(* IEC 61131-3 sources: plcassist-cli/packages/volt-lsp-iec/test-corpus/pro2193/Device/Plc Logic/Application/09 Misc/Library Manager/L_MC4P_RoboticHandling (part 3) *)

(* ---- L_MC4P_PATHREFFROMFILE.fb ---- *)
FUNCTION_BLOCK L_MC4P_PATHREFFROMFILE
VAR_INPUT
	XEXECUTE : BOOL;
	SFILENAME : STRING;
	XABORT : BOOL;
	DWSKIPMASK : DWORD := 0;
	LIBLOCKSEARCHLINENO : LINT := 0;
END_VAR
VAR_OUTPUT
	XDONE : BOOL;
	XBUSY : BOOL;
	XCOMMANDABORTED : BOOL;
	XERROR : BOOL;
	EERRORID : L_IE1P_Error;
	XDECODING : BOOL;
	LILINENODECODED : LINT;
	SLINEDECODED : STRING;
END_VAR
VAR
	LIBLOCKSEARCHLINENO_INT : LINT;
	IFILENO_INT : INT;
	XINTERPRETERHALT_INT : BOOL;
	XMOVEPATHACTIVE_INT : BOOL;
	WACTIVEMFUNCTION_INT : WORD;
	LISOURCELINENO_INT : LINT;
	XABORTACTIVE : BOOL;
	_XDONE : BOOL;
	_XBUSY : BOOL;
	_XCOMMANDABORTED : BOOL;
	_XDECODING : BOOL;
	SFILEADRESS : STRING;
	ITACKEDNUMOFELEMENTSINCYCLE_INT : INT := 0;
	IDECODEMAXNUMOFELEMENTS_INT : INT := 2;
	IDECODEMAXNUMOFELEMENTSFIRSTTIME_INT : INT := 3;
	IDECODENUMOFELEMENTS_INT : INT;
	FB_DECODENCPROGDATA : L_MC1P_StackControlArray := STRUCT(iMaxLegth := GVL_MovePath.gciNumOfPathFiles);
	SCHEADDATA : L_MC4P_AsciiDecoderHeadData;
	RSCACTFILEDATA : REFERENCE TO L_MC4P_AsciiDecoderFileData;
	XHALTATMOS_INT : BOOL := TRUE;
	XIGNOREMCOMMANDS_INT : BOOL;
	XNEWFILE_INT : BOOL;
	LRCIRCLTARGETTOLERANCE_INT : LREAL := 0.1;
	FB_SEMA : L_MC1P_CriticalSection;
	ITAKEELEMENTCNT : INT;
	IADDELEMENTCNT : INT;
	FB_DECODEMOVEDATALOWTASK : L_MC1P_StackControlArray := STRUCT(iMaxLegth := GVL_MovePath.gciNumOfDecodeAsciiData);
	FB_DECODEMOVEDATAMOTIONTASK : L_MC1P_StackControlArray := STRUCT(iMaxLegth := GVL_MovePath.gciNumOfDecodeAsciiData);
	ASCDECODEMOVEDATA_INT : ARRAY [1..GVL_MovePath.gciNumOfDecodeAsciiData] OF L_MC4P_Parameter_MCMove;
	IELEMENINARRAYDECODING : INT;
	FB_DECODEMOVEDATALOWTASK_RESERVE : L_MC1P_StackControlArray := STRUCT(iMaxLegth := GVL_MovePath.gciNumOfDecodeAsciiData_reserve);
	ASCDECODEMOVEDATA_RESERVE : ARRAY [1..GVL_MovePath.gciNumOfDecodeAsciiData_reserve] OF L_MC4P_Parameter_MCMove;
	XERROR_DECODERENDLOOP : BOOL;
	DWTIMEOUTCNT : DWORD := 0;
	DWTIMEOUT : DWORD := 100000;
	XERROR_TIMEOUT : BOOL;
	DWTIMEOUT_MASK : DWORD;
	WTIMEOUTDECODERSTATE : WORD;
	WSTATE : WORD;
	XID1 : BOOL;
	XWID_INT : POINTER TO BOOL := ADR(xId1);
	XSETPATHDATAACTIVE_INT : BOOL;
	XSETPATHDATAACTIVE_OLD : BOOL;
	REQUESTSINFO : DWORD;
	REQUESTSINFO_OLD : DWORD;
	DWRTRIG : DWORD;
	DWFTRIG : DWORD;
	XRESETOUTPUTS : BOOL;
	XERROR_INVALIDSYNCDATA : BOOL;
	BYERRORADRESS : BYTE;
	STERRORADRESSVALUE : STRING;
	XPATHREFABORT : BOOL;
	XDECODEINNEXTTASKCYCLE : BOOL;
	XFBISABORTED : BOOL;
	SFILE_INT : STRING := '';
	XDECODEBUSY_INT : BOOL;
	XDECODEDONE_INT : BOOL;
	XDECODEERROR_INT : BOOL;
	EDECODEEERRORID_INT : L_IE1P_Error;
	DWINTERNALID_INT : DWORD;
	STDECODEERRORLINE : STRING;
	RES : SYSFILE.RTS_IEC_RESULT;
	HFILE : SYSFILE.RTS_IEC_HANDLE;
	UDILENGTHFILE : UDINT;
	XTESTINMOTIONTASK : BOOL := FALSE;
	EXCEPTIONCODE : __SYSTEM.ExceptionCode;
	DWPREDECODERIDLECYCLES : DWORD := 0;
	DWPOSTDECODERIDLECYCLES : DWORD := 0;
	BLOCKSEARCHENABLED : BOOL;
	DATATYPE : WORD;
	DWTIMEOUTMASK : DWORD;
	ENDELEMENT : POINTER TO L_MC4P_Parameter_MCMove;
	ENDIDX : INT;
	POSTDECODERIDLECYCLES : DWORD;
	PREDECODERIDLECYCLES : DWORD;
	SETCIRCTARGETTOLERANCE : LREAL;
	SIZE : UDINT;
	STARTELEMENT : POINTER TO L_MC4P_Parameter_MCMove;
	STARTIDX : INT;
	STERRORCOMMAND : STRING;
	TAKEELEMENT : POINTER TO L_MC4P_Parameter_MCMove;
	XDECODEINMOTIONTASK : BOOL;
	XHALTATMOS : BOOL;
	XIGNOREMCOMMANDS : BOOL;
	XINTERPRETERHALT : BOOL;
END_VAR
END_FUNCTION_BLOCK

METHOD ABORTFB
END_METHOD

METHOD CALL_ALLOCPOINTADR
END_METHOD

METHOD CALL_ERRORHANDLER
END_METHOD

METHOD CALL_FBMETHODS
END_METHOD

METHOD CALL_OUTPUT
END_METHOD

METHOD CALL_REQUESTS_EXT
END_METHOD

METHOD CALL_RESETCOMMANDS
END_METHOD

METHOD CALL_RESETOUTPUT
END_METHOD

METHOD CALL_RESETSTATUS
END_METHOD

METHOD CALL_STATEMACHINE
END_METHOD

METHOD CALL_SYNCDECODEMOVEDATA
END_METHOD

METHOD FUN_DECODEAUX : BOOL
VAR_IN_OUT
	STADRESSVALUE : STRING(255);
	SCDECODEHEADDATA : L_MC4P_AsciiDecoderHeadData;
END_VAR
END_METHOD

METHOD FUN_DECODEADRESS : BOOL
VAR_OUTPUT
	XERROR : BOOL;
	EERRORID : L_IE1P_Error;
END_VAR
VAR_IN_OUT
	BYADRESS : BYTE;
	STADRESSVALUE : STRING(255);
	SCDECODEHEADDATA : L_MC4P_AsciiDecoderHeadData;
END_VAR
END_METHOD

METHOD FUN_DECODEG : BOOL
VAR_IN_OUT
	LIADRESSVALUE : LINT;
	SCDECODEHEADDATA : L_MC4P_AsciiDecoderHeadData;
END_VAR
END_METHOD

METHOD FUN_DECODEGOTO : BOOL
VAR_OUTPUT
	XERROR : BOOL;
	EERRORID : L_IE1P_Error;
END_VAR
VAR_IN_OUT
	STADRESSVALUE : STRING(255);
	SCDECODEHEADDATA : L_MC4P_AsciiDecoderHeadData;
END_VAR
END_METHOD

METHOD FUN_DECODEH : BOOL
VAR_IN_OUT
	STADRESSVALUE : STRING(255);
	SCDECODEHEADDATA : L_MC4P_AsciiDecoderHeadData;
	XERROR : BOOL;
	EERRORID : L_IE1P_Error;
END_VAR
END_METHOD

METHOD FUN_DECODEI : BOOL
VAR_IN_OUT
	STADRESSVALUE : STRING(255);
	SCDECODEHEADDATA : L_MC4P_AsciiDecoderHeadData;
END_VAR
END_METHOD

METHOD FUN_DECODEIFCASE : BOOL
VAR_INPUT
	STLINE : STRING(255);
END_VAR
VAR_OUTPUT
	XERROR : BOOL;
	EERRORID : L_IE1P_Error;
END_VAR
VAR_IN_OUT
	SCDECODEHEADDATA : L_MC4P_AsciiDecoderHeadData;
END_VAR
END_METHOD

METHOD FUN_DECODEL : BOOL
VAR_IN_OUT
	STADRESSVALUE : STRING(255);
	SCDECODEHEADDATA : L_MC4P_AsciiDecoderHeadData;
	XERROR : BOOL;
	EERRORID : L_IE1P_Error;
END_VAR
END_METHOD

METHOD FUN_DECODELINE : BOOL
VAR_OUTPUT
	XGETNEXTSOURCELINE : BOOL;
	XELEMENTDECODED : BOOL;
	XERROR : BOOL;
	EERRORID : L_IE1P_Error;
END_VAR
VAR_IN_OUT
	SCDECODEHEADDATA : L_MC4P_AsciiDecoderHeadData;
	SCDECODEMOVEDATA : L_MC4P_Parameter_MCMove;
END_VAR
END_METHOD

METHOD FUN_DECODEM : BOOL
VAR_IN_OUT
	LIADRESSVALUE : LINT;
	SCDECODEHEADDATA : L_MC4P_AsciiDecoderHeadData;
	XERROR : BOOL;
	EERRORID : L_IE1P_Error;
END_VAR
END_METHOD

METHOD FUN_DECODEN : BOOL
VAR_IN_OUT
	STADRESSVALUE : STRING(255);
	SCDECODEHEADDATA : L_MC4P_AsciiDecoderHeadData;
END_VAR
END_METHOD

METHOD FUN_DECODEO : BOOL
VAR_IN_OUT
	STADRESSVALUE : STRING(255);
	SCDECODEHEADDATA : L_MC4P_AsciiDecoderHeadData;
	XERROR : BOOL;
	EERRORID : L_IE1P_Error;
END_VAR
END_METHOD

METHOD FUN_DECODEP : BOOL
VAR_IN_OUT
	STADRESSVALUE : STRING(255);
	SCDECODEHEADDATA : L_MC4P_AsciiDecoderHeadData;
END_VAR
END_METHOD

METHOD FUN_DELETECOMMENTS : BOOL
VAR_OUTPUT
	STCOMMENT : STRING;
	ILINESIZE : INT;
END_VAR
VAR_IN_OUT
	STLINE : STRING(255);
END_VAR
END_METHOD

METHOD FUN_DELETECOMMENTS_TYPE1 : BOOL
VAR_IN_OUT
	STLINE : STRING(255);
	STCOMMENT : STRING;
	ICOMMENTPOS : INT;
END_VAR
END_METHOD

METHOD FUN_DELETECOMMENTS_TYPE2 : BOOL
VAR_INPUT
	ICOMMENTTYPE : INT;
END_VAR
VAR_IN_OUT
	STLINE : STRING(255);
	STCOMMENT : STRING;
END_VAR
END_METHOD

METHOD FUN_FINDJUMPTARB : BOOL
VAR_INPUT
	LIJUMPTARGET : LINT;
	UDIFILELENGTH : UDINT;
	UDIPOS : UDINT;
	UDIPOSSTART : UDINT;
END_VAR
VAR_OUTPUT
	UDITARLINEPOS : UDINT;
	XERROR : BOOL;
	EERRORID : L_IE1P_Error;
END_VAR
END_METHOD

METHOD FUN_FINDJUMPTARF : BOOL
VAR_INPUT
	LIJUMPTARGET : LINT;
	UDIFILELENGTH : UDINT;
	UDIPOS : UDINT;
END_VAR
VAR_OUTPUT
	UDITARLINEPOS : UDINT;
	XERROR : BOOL;
	EERRORID : L_IE1P_Error;
END_VAR
END_METHOD

METHOD FUN_GOTO : BOOL
VAR_OUTPUT
	XERROR : BOOL;
	EERRORID : L_IE1P_Error;
END_VAR
VAR_IN_OUT
	SCDECODEHEADDATA : L_MC4P_AsciiDecoderHeadData;
	STLINE : STRING(255);
END_VAR
END_METHOD

METHOD FUN_GETADRESS : BOOL
VAR_OUTPUT
	ILINESIZE : INT;
	BYADRESS : BYTE;
	SADRESSVALUE : STRING;
END_VAR
VAR_IN_OUT
	STLINE : STRING(255);
END_VAR
END_METHOD

METHOD FUN_ISALPHACHAR : BOOL
VAR_INPUT
	BYCHAR : BYTE;
END_VAR
END_METHOD

METHOD FUN_READLINE : L_IE1P_Error
VAR_INPUT
	UDIPOSIN : UDINT;
	XEXITCLOSEFILE : BOOL;
	XFINDSTARTCOMAND : BOOL;
END_VAR
VAR_OUTPUT
	UDIPOSOUT : UDINT;
	ILINESIZE : INT;
	IPOSLF : INT;
	IPOSNL : INT;
	UDIRESULTFILEOPEN : UDINT;
	UDIRESULTREADSTRING : UDINT;
	XENDOFFILE : BOOL;
	XLASTLINE : BOOL;
	XSTART : BOOL;
END_VAR
VAR_IN_OUT
	HFILE : SYSFILE.RTS_IEC_HANDLE;
	RES : SYSFILE.RTS_IEC_ResULT;
	STLINE : STRING(255);
END_VAR
END_METHOD

METHOD FUN_READLINEBACK : BOOL
VAR_INPUT
	UDIPOSIN : UDINT;
	XEXITCLOSEFILE : BOOL;
	UDIPOSSTART : UDINT := 0;
END_VAR
VAR_OUTPUT
	UDIPOSOUT : UDINT;
	ILINESIZE : INT;
	UDIRESULTFILEOPEN : UDINT;
	XSTARTOFFILE : BOOL;
END_VAR
VAR_IN_OUT
	HFILE : SYSFILE.RTS_IEC_HANDLE;
	RES : SYSFILE.RTS_IEC_ResULT;
	STLINE : STRING(255);
END_VAR
END_METHOD

METHOD FUN_REPLACEVAR : BOOL
VAR_IN_OUT
	STVALUE : STRING(255);
END_VAR
END_METHOD

METHOD FUN_STRING_PLCVARIABLE_TO_LINT : BOOL
VAR_INPUT
	STVALUE : STRING(255);
END_VAR
VAR_OUTPUT
	LIVALUE : LINT;
END_VAR
END_METHOD

METHOD FUN_STRING_PLCVARIABLE_TO_LREAL : BOOL
VAR_INPUT
	STVALUE : STRING(255);
END_VAR
VAR_OUTPUT
	LRVALUE : LREAL;
END_VAR
END_METHOD

METHOD FUN_STRING_TO_LINT : BOOL
VAR_INPUT
	STVALUE : STRING;
	XVARALLOWED : BOOL;
END_VAR
VAR_OUTPUT
	LIVALUE : LINT;
END_VAR
END_METHOD

METHOD FUN_STRING_TO_LREAL : BOOL
VAR_INPUT
	STVALUE : STRING(255);
END_VAR
VAR_OUTPUT
	LRVALUE : LREAL;
END_VAR
END_METHOD

METHOD FUN_SHUNTINGYARD : BOOL
VAR_INPUT
	STVALUE : STRING(255);
END_VAR
VAR_OUTPUT
	SCVALUE : L_UBUP_Variable;
END_VAR
END_METHOD

METHOD CALL_DECODER
END_METHOD

METHOD CALL_DECODER_READASCIIFILE
END_METHOD

METHOD EXECUTEFREERUNTASK
END_METHOD

METHOD FUN_CLOSEFILE
END_METHOD

METHOD INIT_HEADDATA
VAR_IN_OUT
	SCDECODEHEADDATA : L_MC4P_AsciiDecoderHeadData;
END_VAR
END_METHOD

METHOD MAIN
END_METHOD

METHOD GETID : __XWORD
END_METHOD

METHOD GETPATHDATA : ARRAY [1..GVL_MovePath.gciNumOfDecodeAsciiData] OF POINTER TO L_MC4P_Parameter_MCMove
END_METHOD

METHOD GETPATHDATAACTIVE : BOOL
END_METHOD

METHOD GETSTATUS : DWORD
END_METHOD

METHOD SETABORT
END_METHOD

METHOD SETACTIVEMFUNCTION
VAR_INPUT
	WACTIVEMFUNCTION : WORD;
END_VAR
END_METHOD

METHOD SETMOVEPATHACTIVE
VAR_INPUT
	XMOVEPATHACTIVE : BOOL;
END_VAR
END_METHOD

METHOD SETPATHDATAACTIVE
VAR_INPUT
	XPATHDATAACTIVE : BOOL;
END_VAR
END_METHOD

METHOD CALL_INIT
END_METHOD

METHOD CALL_S000_CYCLIC
END_METHOD

METHOD ABORT : UDINT
END_METHOD

METHOD EXECUTE : UDINT
END_METHOD

(* ---- L_MC4P_PATHREFMONITOR.fb ---- *)
FUNCTION_BLOCK L_MC4P_PATHREFMONITOR
VAR_INPUT
	XEXECUTE : BOOL;
	XABORT : BOOL;
	ITFPATHREF : MC_PATH_REF;
	SCSKIP : L_MC4P_SkipGCode;
	ASCDATA : POINTER TO L_MC4P_PathRefMonitorData;
END_VAR
VAR_OUTPUT
	XDONE : BOOL;
	XBUSY : BOOL;
	XCOMMANDABORTED : BOOL;
	XERROR : BOOL;
	EERRORID : L_IE1P_Error;
	UDINEWESTELEMENT : UDINT;
	UDIELEMENTCOUNT : UDINT;
END_VAR
VAR
	_ITFPATHREF : MC_PATH_REF;
	_UDISTARTIDX : UDINT;
	_UDIENDIDX : UDINT;
	_UDIREADIDX : UDINT;
	_UDILOWER : UDINT;
	_UDIUPPER : UDINT;
	_UDISIZE : UDINT;
	_DWSTATUS : DWORD;
	_XREINIT : BOOL := FALSE;
	_XDATADIALOG : BOOL := FALSE;
	_UDIVISUARRIDX : UDINT := 0;
	_PSCDATAARR : POINTER TO L_MC4P_PathRefMonitorData;
	_PSCDATAVISU : POINTER TO L_MC4P_PathRefMonitorData;
	_SCDATAINITIAL : L_MC4P_PathRefMonitorData;
	_ISKIPVIEWFRAME : INT := 0;
	_MODEL : L_UBUP_BehaviourModel_ETrigA;
END_VAR
END_FUNCTION_BLOCK

METHOD MAPOUTPUTS
END_METHOD

METHOD CYCLICACTION
VAR_INPUT
	ITFTIMINGCONTROLLER : L_UBUP.L_UBUP_ITimingController;
END_VAR
VAR_OUTPUT
	XCOMPLETE : BOOL;
	XABORT : BOOL;
	IERRORID : INT;
END_VAR
END_METHOD

METHOD FINALIZEACTION
VAR_INPUT
	XABORTPROPOSED : BOOL;
	IERRORIDPROPOSED : INT;
END_VAR
VAR_OUTPUT
	XCOMPLETE : BOOL;
	XABORT : BOOL;
	IERRORID : INT;
END_VAR
END_METHOD

METHOD RESETACTION
VAR_OUTPUT
	XCOMPLETE : BOOL;
END_VAR
END_METHOD

METHOD STARTACTION
VAR_OUTPUT
	XCOMPLETE : BOOL;
	IERRORID : INT;
END_VAR
END_METHOD

METHOD FB_INIT : BOOL
VAR_INPUT
	BINITRETAINS : BOOL;
	BINCOPYCODE : BOOL;
END_VAR
END_METHOD

METHOD APPENDDATASET : BOOL
VAR_INPUT
	PMCMOVE : POINTER TO L_MC4P_Parameter_MCMove;
END_VAR
END_METHOD

METHOD SKIP : BOOL
VAR_INPUT
	PMCMOVE : POINTER TO L_MC4P_Parameter_MCMove;
END_VAR
END_METHOD

(* ---- L_MC4P_PICKANDPLACEMEMORY.fb ---- *)
FUNCTION_BLOCK L_MC4P_PICKANDPLACEMEMORY
VAR_INPUT
	FB_SEMAMOVEFBS : L_MC1P_CriticalSection;
	AMC_MOVELINREL : ARRAY [1..3] OF L_MC4P_MoveLinearRelative_Internal;
	AFB_MOVEELLIPTICAL : ARRAY [1..3] OF L_MC4P_MoveEllipticalAbsolutePnP_Internal;
	AFB_MOVESPLINE : ARRAY [1..3] OF L_MC4P_MoveSplinePnP_Internal;
	AMC_MOVELINABS1 : ARRAY [1..10] OF L_MC4P_MoveLinearAbsolute_Internal;
	AMC_MOVELINABS2 : ARRAY [1..10] OF L_MC4P_MoveLinearAbsolute_Internal;
	AMC_MOVELINABS3 : ARRAY [1..10] OF L_MC4P_MoveLinearAbsolute_Internal;
	AMC_MOVELINABS4 : ARRAY [1..3] OF L_MC4P_MoveLinearAbsolute_Internal;
	AMC_MOVELINABS5 : ARRAY [1..2] OF L_MC4P_MoveLinearAbsolute_Internal;
	AMC_MOVEDIRABS1 : ARRAY [1..10] OF L_MC4P_MoveDirectAbsolute_Internal;
	AMC_MOVEDIRABS2 : ARRAY [1..10] OF L_MC4P_MoveDirectAbsolute_Internal;
	AMC_MOVEDIRREL : ARRAY [1..1] OF L_MC4P_MoveDirectRelative_Internal;
	AFB_GROUPWAITTIME : ARRAY [1..3] OF L_MC4P_GroupWaitTime_Internal;
	ASCPROFILEPARMEM : ARRAY [1..10] OF ARRAY [1..10] OF L_MC4P_scPickAndPlaceProfileParState;
	ASCPROFILETIMEFROMCVTARGET : ARRAY [1..16] OF ARRAY [0..10] OF L_MC4P_MeasuredProfileTime;
	AIRINGMEMPROFILETIME : ARRAY [1..16] OF ARRAY [1..2] OF INT;
	FB_SEMA : L_MC1P_CriticalSection;
	CONVEYORBELTVIRTUAL : ARRAY [1..2] OF AXIS_REF := [STRUCT(UsedAsInternalAxisInstance := TRUE), STRUCT(UsedAsInternalAxisInstance := TRUE)];
END_VAR
END_FUNCTION_BLOCK

(* ---- L_MC4P_PREPAREPATH.fb ---- *)
FUNCTION_BLOCK L_MC4P_PREPAREPATH EXTENDS L_MC4P_Template_KIN
VAR_INPUT
	PLIST : POINTER TO L_MC4P_PathDataList;
	PPATHELEMENT : POINTER TO L_MC4P_PathElement;
	ALRSTARTPOS : ARRAY [1..12] OF LREAL;
	PAXESGROUP : POINTER TO AXES_GROUP_KIN;
	XINITSTATEMACHINE : BOOL;
	PCORRESPONDINGFB : POINTER TO L_MC4P_MoveContPath;
	XCHECKWORKSPACE : BOOL := TRUE;
	UDICHECKWORKSPACESTEPS : UDINT := 5;
END_VAR
VAR_OUTPUT
	XERROR : BOOL := FALSE;
	ERRORID : L_IE1P_Error;
	DWINTERNALERRORID : DWORD;
END_VAR
VAR
	SCERROR : L_MC4P_ErrorStruct;
	XNOBLENDINGERRORS : BOOL := TRUE;
	XDOPREPARE : BOOL := FALSE;
	PLISTELEMENT : POINTER TO L_MC4P_ListElement;
	PLISTELEMENT_PREVIOUS : POINTER TO L_MC4P_ListElement;
	PLISTELEMENTSTART : POINTER TO L_MC4P_ListElement;
	PLISTELEMENTEND : POINTER TO L_MC4P_ListElement;
	PLISTELEMENT_IDENTPTPTYPE : POINTER TO L_MC4P_ListElement;
	PLISTELEMENT_CALCPTPPROFILE : POINTER TO L_MC4P_ListElement;
	WSTEP : WORD := 0;
	PTP_PREPSTATE : L_MC4P_PTPPrepStates;
	BIDENTTMAX_INIT : BOOL;
	BIDENTPTPTYPE_INIT : BOOL;
	BCALCPTPPROFILE_INIT : BOOL;
	ACHSE : UINT;
	CNTCYCLESPREPAREPATH : UINT;
	CNTCYCLESPREPAREPATHMAX : UINT := 500;
	BYAUXAXISSEQCOUNT : BYTE;
	PLISTELEMENTAUXSEQSTART : ARRAY [1..6] OF POINTER TO L_MC4P_ListElement;
	PLISTELEMENTAUXSEQEND : ARRAY [1..6] OF POINTER TO L_MC4P_ListElement;
	XRECALCPROFILES : BOOL;
	XAUXAXISACTIVNEWSET : BOOL;
	PTESTAUX : POINTER TO L_MC4P_ListElement;
	XFOUND : BOOL;
	LRTIMEELEMENT : LREAL;
	LRJERKDEC : LREAL;
	DWIPOSTATE : DWORD;
	LRTIMELIST : LREAL;
	LRTIMEIPO : LREAL;
	LRTIMEREST : LREAL;
	LRTIMETOCUT : LREAL;
	LRTIMEACCZERO : LREAL;
	LRSTARTACC : LREAL;
	LRSTARTVEL : LREAL;
	LRSTARTPOS : LREAL;
	LRENDACC : LREAL;
	LRENDVEL : LREAL;
	LRENDPOS : LREAL;
	DWBOTHDIRECTIONS : DWORD := 3;
	SCPROFILEPARAMETER : L_MC1P_ProfileParameter;
	SCPROFILEDATA : L_MC1P_ProfileData;
	PLISTELEMENTTMP : POINTER TO L_MC4P_ListElement;
	WCPP_ABC_STEP : WORD;
	WCPPSTEP : WORD;
	LRVIN_ORIGINAL : LREAL;
	LRVOUT_ORIGINAL : LREAL;
	XDOPROFILECHECK : BOOL := FALSE;
	WDOPREPARECOUNTER : WORD;
	WDOPREPARECOUNTERMAX : WORD := 1;
	WLDE_MODE : WORD := 2;
	LRANGULARTOLERANCE_LDC : LREAL := 0.1;
	LRMAXACCDIFF_LDC : LREAL := 0.0;
	LRACCREDFACTOR : LREAL := 0.1;
	TIMESTART : ULINT;
	TIMEEND : ULINT;
	AXTAKETIMESTAMP : ARRAY [0..20] OF BOOL;
	ULIPREPPATHTIME : ARRAY [0..20] OF ULINT;
	DWSCHELLINGWORKAROUNDCOUNTER : DWORD := 0;
	DIRESETBLENDINGSEGMENTNO : DINT := 0;
	DIBLENDINGSEGMENTNORESETTED : DINT := 0;
	XBLENDINGALWAYSSHORTESTWAY : BOOL := FALSE;
	XENABLECORRLDS00042356 : BOOL := TRUE;
	SCSP : L_MC4P_CyclicData;
	LRPERCLENGTHDELTA : LREAL := 0.1;
	LRFACTOR : LREAL := (1 / (1.0 - (0.1 * lrPercLengthDelta)));
END_VAR
END_FUNCTION_BLOCK

METHOD ACTIVATESEGMENT
VAR_INPUT
	PLISTELEMENT : POINTER TO L_MC4P_ListElement;
END_VAR
END_METHOD

METHOD AUXAXISCALCMAINPATHLENGTH : BOOL
VAR_INPUT
	PLISTELEMENT : POINTER TO L_MC4P_ListElement;
	IDX : INT;
END_VAR
VAR_OUTPUT
	LRMAINAXPATH : LREAL;
	PLISTELEMENTAUXSEQSTART : POINTER TO L_MC4P_ListElement;
END_VAR
END_METHOD

METHOD AUXAXISCALCMAINTIME : BOOL
VAR_INPUT
	PLISTELEMENT : POINTER TO L_MC4P_ListElement;
	IDX : INT;
END_VAR
VAR_OUTPUT
	LRMAINTIMECOMPLETE : LREAL;
	LRMAINAXPATH : LREAL;
	PLISTELEMENTAUXSEQSTART : POINTER TO L_MC4P_ListElement;
END_VAR
END_METHOD

METHOD AUXAXISLIMITMAINAXIS
VAR_INPUT
	PLISTELEMENT : POINTER TO L_MC4P_ListElement;
END_VAR
VAR_OUTPUT
	XRECALCPROFILES : BOOL := FALSE;
END_VAR
END_METHOD

METHOD AUXAXISPREPARE
VAR_INPUT
	PLISTELEMENT : POINTER TO L_MC4P_ListElement;
END_VAR
VAR_OUTPUT
	XRECALCPROFILES : BOOL := FALSE;
END_VAR
END_METHOD

METHOD CALCULATEORIPATH
VAR_INPUT
	PLISTELEMENTDATA : POINTER TO L_MC4P_ListElementData;
END_VAR
END_METHOD

METHOD CALCULATEPTPTARGET
VAR_INPUT
	PLISTELEMENTDATA : POINTER TO L_MC4P_ListElementData;
END_VAR
END_METHOD

METHOD CALCULATEPATHPOLYNOM
VAR_INPUT
	PLISTELEMENT : POINTER TO L_MC4P_ListElement;
END_VAR
END_METHOD

METHOD CALCULATEPROFILEABC
VAR_INPUT
	PLISTELEMENT : POINTER TO L_MC4P_ListElement;
END_VAR
VAR_OUTPUT
	XSTEPBACK : BOOL;
END_VAR
END_METHOD

METHOD CALCULATEPROFILEPOLYNOM
VAR_INPUT
	PLISTELEMENT : POINTER TO L_MC4P_ListElement;
END_VAR
END_METHOD

METHOD CREATERESETBLENDINGLOG
END_METHOD

METHOD DETERMINEBLENDINGDIRECTION : BOOL
VAR_INPUT
	PREVIOUS : POINTER TO L_MC4P_ListElementData;
	BLENDING : POINTER TO L_MC4P_ListElementData;
	NEXT : POINTER TO L_MC4P_ListElementData;
END_VAR
END_METHOD

METHOD INTERPRETER
VAR_INPUT
	PPATHELEMENT : POINTER TO L_MC4P_PathElement;
END_VAR
VAR_IN_OUT
	PLIST : POINTER TO L_MC4P_PathDataList;
END_VAR
END_METHOD

METHOD LIMITDYNAMICSCOMBINE
VAR_INPUT
	PLISTELEMENT : POINTER TO L_MC4P_ListElement;
END_VAR
END_METHOD

METHOD LIMITDYNAMICSCORNER
VAR_INPUT
	PLISTELEMENT : POINTER TO L_MC4P_ListElement;
END_VAR
END_METHOD

METHOD LIMITDYNAMICSELEMENTS
VAR_INPUT
	PLISTELEMENT : POINTER TO L_MC4P_ListElement;
END_VAR
END_METHOD

METHOD LIMITDYNAMICSPATHLENGTH
VAR_INPUT
	PLISTELEMENTSTART : POINTER TO L_MC4P_ListElement;
	PLISTELEMENTEND : POINTER TO L_MC4P_ListElement;
END_VAR
END_METHOD

METHOD LIMITDYNAMICSPATHLENGTH_KART
VAR_INPUT
	PLISTELEMENTSTART : POINTER TO L_MC4P_ListElement;
	PLISTELEMENTEND : POINTER TO L_MC4P_ListElement;
END_VAR
END_METHOD

METHOD PREPAREPTPPROFILES
VAR_INPUT
	PLISTELEMENTSTART : POINTER TO L_MC4P_ListElement;
	PLISTELEMENTEND : POINTER TO L_MC4P_ListElement;
END_VAR
END_METHOD

METHOD PREPAREPTPPROFILES_CALCPTPPROFILE
VAR_INPUT
	PLISTELEMENTSTART : POINTER TO L_MC4P_ListElement;
	PLISTELEMENTEND : POINTER TO L_MC4P_ListElement;
END_VAR
VAR_OUTPUT
	XRETURN : BOOL;
END_VAR
END_METHOD

METHOD PREPAREPTPPROFILES_IDENTPTPTYPE
VAR_INPUT
	PLISTELEMENTSTART : POINTER TO L_MC4P_ListElement;
	PLISTELEMENTEND : POINTER TO L_MC4P_ListElement;
END_VAR
VAR_OUTPUT
	XRETURN : BOOL;
END_VAR
END_METHOD

METHOD PREPAREPTPPROFILES_IDENTTMAX
VAR_INPUT
	PLISTELEMENTSTART : POINTER TO L_MC4P_ListElement;
	PLISTELEMENTEND : POINTER TO L_MC4P_ListElement;
END_VAR
VAR_OUTPUT
	XRETURN : BOOL;
END_VAR
END_METHOD

METHOD PREPAREPTPPROFILES_QUITPREP
VAR_INPUT
	PLISTELEMENTSTART : POINTER TO L_MC4P_ListElement;
	PLISTELEMENTEND : POINTER TO L_MC4P_ListElement;
END_VAR
END_METHOD

METHOD RAISESWLIMITERROR : L_IE1P_Error
VAR_INPUT
	PLISTELEMENT : POINTER TO L_MC4P_ListElement;
	IDX : DINT;
END_VAR
END_METHOD

METHOD RESETPATHANDRESTART
END_METHOD

METHOD RESETPATHPREPARATION
END_METHOD

METHOD SMOOTHPATH
VAR_INPUT
	PLISTELEMENT : POINTER TO L_MC4P_ListElement;
END_VAR
END_METHOD

METHOD STRETCHPROFILETOTIME
VAR_INPUT
	PROFILEDATA_ACT : L_MC1P_ProfileData;
	PARAM_ACT : L_MC1P_ProfileParameter;
	T_DESIRED : LREAL;
END_VAR
VAR_OUTPUT
	PROFILEDATA_NEW : L_MC1P_ProfileData;
	PARAM_NEW : L_MC1P_ProfileParameter;
END_VAR
END_METHOD

METHOD CALC_RAST2VEL_TRAPONLY
VAR_INPUT
	POS_IN : LREAL;
	POS_OUT : LREAL;
	JERK : LREAL;
	AMAX : LREAL;
	T_DESIRED : LREAL;
END_VAR
VAR_IN_OUT
	SCPROFILEDATA : L_MC1P_ProfileData;
END_VAR
END_METHOD

METHOD CALC_RAST2VEL_TRIONLY
VAR_INPUT
	POS_IN : LREAL;
	POS_OUT : LREAL;
	JERK : LREAL;
	T_DESIRED : LREAL;
END_VAR
VAR_IN_OUT
	SCPROFILEDATA : L_MC1P_ProfileData;
END_VAR
END_METHOD

METHOD CALC_REDVMAX
VAR_INPUT
	ACT : POINTER TO L_MC4P_ListElementData;
	ACHSE : UINT;
	T_MAX_ACT : LREAL;
END_VAR
END_METHOD

METHOD CALC_VEL2RAST_TRAPONLY
VAR_INPUT
	POS_IN : LREAL;
	POS_OUT : LREAL;
	JERK : LREAL;
	V_IN : LREAL;
	AMAX : LREAL;
	T_DESIRED : LREAL;
END_VAR
VAR_IN_OUT
	SCPROFILEDATA : L_MC1P_ProfileData;
END_VAR
END_METHOD

METHOD CALC_VEL2RAST_TRIONLY
VAR_INPUT
	POS_IN : LREAL;
	POS_OUT : LREAL;
	JERK : LREAL;
	V_IN : LREAL;
	V_OUT : LREAL;
	AMAX : LREAL;
	T_DESIRED : LREAL;
END_VAR
VAR_IN_OUT
	SCPROFILEDATA : L_MC1P_ProfileData;
END_VAR
END_METHOD

METHOD CREATEABCELEMENTS
VAR_INPUT
	PLISTELEMENTCUT : POINTER TO L_MC4P_ListElement;
END_VAR
VAR_OUTPUT
	PLISTELEMENTCUT_1A : POINTER TO L_MC4P_ListElement;
	PLISTELEMENTCUT_1B : POINTER TO L_MC4P_ListElement;
	PLISTELEMENTCUT_1C : POINTER TO L_MC4P_ListElement;
	PLISTELEMENTCUT_2B : POINTER TO L_MC4P_ListElement;
	PLISTELEMENTCUT_2C : POINTER TO L_MC4P_ListElement;
	PNEW : POINTER TO L_MC4P_ListElement;
	PLEFT : POINTER TO L_MC4P_ListElement;
END_VAR
END_METHOD

METHOD IDENTCUTELEMENT
VAR_IN_OUT
	PLISTELEMENTCUT : POINTER TO L_MC4P_ListElement;
END_VAR
END_METHOD

METHOD LOOKAHEAD_CLEANUP
END_METHOD

METHOD LOOKAHEAD_PREPARE
END_METHOD

METHOD MODIFYABCELEMENTS
VAR_INPUT
	PLISTELEMENTCUT : POINTER TO L_MC4P_ListElement;
END_VAR
VAR_IN_OUT
	PLISTELEMENTCUT_1A : POINTER TO L_MC4P_ListElement;
	PLISTELEMENTCUT_1B : POINTER TO L_MC4P_ListElement;
	PLISTELEMENTCUT_1C : POINTER TO L_MC4P_ListElement;
END_VAR
END_METHOD

METHOD CALCMAXVELOUT : LREAL
VAR_INPUT
	LRJERK : LREAL;
	LRAMAX : LREAL;
	LRDIST : LREAL;
	LRVIN : LREAL;
END_VAR
END_METHOD

METHOD INITGEOOBJECT
VAR_INPUT
	PLISTELEMENT : POINTER TO L_MC4P_ListElement;
END_VAR
VAR_OUTPUT
	SCERROR : L_MC4P_ErrorStruct;
END_VAR
END_METHOD

METHOD CHECKWORKSPACE
VAR_INPUT
	PLISTELEMENT : POINTER TO L_MC4P_ListElement;
END_VAR
END_METHOD

METHOD CHECKWORKSPACEDOT
VAR_INPUT
	PLISTELEMENT : POINTER TO L_MC4P_ListElement;
	LRPERCLENGTH : LREAL;
	LRLENGTH : LREAL;
	SCTRAFOINFO_SW : REFERENCE TO L_MC4P_TrafoInfo;
	SCERROR : REFERENCE TO L_MC4P_ErrorStruct;
END_VAR
END_METHOD

(* ---- L_MC4P_READBOOLPARAMETER.fb ---- *)
FUNCTION_BLOCK L_MC4P_READBOOLPARAMETER EXTENDS L_MC4P_Template_AG_KIN
VAR_INPUT
	XENABLE : BOOL;
	DIPARAMETERNUMBER : DINT;
END_VAR
VAR_OUTPUT
	XVALID : BOOL;
	XBUSY : BOOL;
	XERROR : BOOL;
	EERRORID : L_IE1P_Error;
	XVALUE : BOOL;
END_VAR
VAR
	XENABLEOLD : BOOL := FALSE;
END_VAR
END_FUNCTION_BLOCK

METHOD FB_RESET : BOOL
END_METHOD

(* ---- L_MC4P_READPARAMETER.fb ---- *)
FUNCTION_BLOCK L_MC4P_READPARAMETER EXTENDS L_MC4P_Template_AG_KIN
VAR_INPUT
	XENABLE : BOOL;
	DIPARAMETERNUMBER : DINT;
END_VAR
VAR_OUTPUT
	XVALID : BOOL;
	XBUSY : BOOL;
	XERROR : BOOL;
	EERRORID : L_IE1P_Error;
	LRVALUE : LREAL;
END_VAR
VAR
	XENABLEOLD : BOOL := FALSE;
END_VAR
END_FUNCTION_BLOCK

METHOD FB_RESET : BOOL
END_METHOD

(* ---- L_MC4P_SETACTIVETOOL.fb ---- *)
FUNCTION_BLOCK L_MC4P_SETACTIVETOOL EXTENDS L_MC4P_Template_AG_KIN
VAR_INPUT
	XEXECUTE : BOOL;
	ETOOLSYSTEM : L_MC4P_ToolSystem;
END_VAR
VAR_OUTPUT
	XDONE : BOOL;
	XBUSY : BOOL;
	XERROR : BOOL;
	EERRORID : L_IE1P_Error := L_IE1P_Error.NoError;
END_VAR
VAR
	XEXECUTEOLD : BOOL;
	XRESETOUTPUT : BOOL;
END_VAR
END_FUNCTION_BLOCK

(* ---- L_MC4P_SETTOOLTRANSFORM.fb ---- *)
FUNCTION_BLOCK L_MC4P_SETTOOLTRANSFORM EXTENDS L_MC4P_Template_AG_KIN
VAR_INPUT
	XEXECUTE : BOOL;
	SCTOOLPARAMETER : L_MC4P_TOOL_REF;
	ETOOLSYSTEM : L_MC4P_ToolSystem;
END_VAR
VAR_OUTPUT
	XDONE : BOOL;
	XBUSY : BOOL;
	XERROR : BOOL;
	EERRORID : L_IE1P_Error := L_IE1P_Error.NoError;
END_VAR
VAR
	PTOOL : POINTER TO L_MC4P_ToolTrafo;
	XEXECUTEOLD : BOOL;
	XRESETOUTPUT : BOOL;
	AXPARACCESSIBLE : ARRAY [1..7] OF BOOL;
	IDX : DINT;
	XINTERNALTESTMODE : BOOL := FALSE;
	INTERNALTESTMODE : BOOL;
END_VAR
END_FUNCTION_BLOCK

(* ---- L_MC4P_SETVALUEFILTER.fb ---- *)
FUNCTION_BLOCK L_MC4P_SETVALUEFILTER EXTENDS L_UBUP_MemoryProvider
VAR_INPUT
	XENABLE : BOOL;
	EFILTERMODE : L_MC4P_SetValueFilterMode := L_MC4P_SetValueFilterMode.EqualySpaced;
	UIFILTERTIME : UINT;
	LRSETPOSIN : LREAL;
	LRSETVELIN : LREAL;
	LRSETACCIN : LREAL;
	LRSETPOSINITIAL : LREAL;
	ETRAVERSINGRANGE : L_MC1P_TraversingRange := L_MC1P_TraversingRange.Limited;
	LRCYCLELENGTH : LREAL;
	LRINVCYCLELENGTH : LREAL;
END_VAR
VAR_OUTPUT
	XBUSY : BOOL;
	XACTIVE : BOOL;
	XERROR : BOOL;
	EERRORID : L_IE1P.L_IE1P_Error;
	DWINTERNALID : DWORD;
	LRSETPOSOUT : LREAL;
	LRSETVELOUT : LREAL;
	LRSETACCOUT : LREAL;
	LRACTFILTERDELAY : LREAL;
END_VAR
VAR
	LRTASKCYCLE : LREAL := -1;
	XENABLE_R : R_Trig;
	AMEM : ARRAY [1..4] OF ARRAY [1..cuiFilterSizeMax] OF LREAL;
	FB_AVG : L_USPP_AverageFilterRecursive;
	CUIFILTERSIZEMAX : UINT := 501;
	XRECURSIVE : BOOL := TRUE;
	PTR : POINTER TO BYTE;
	SIZE : UDINT;
END_VAR
END_FUNCTION_BLOCK

(* ---- L_MC4P_SIMPLETRANSFORMATION.fb ---- *)
FUNCTION_BLOCK L_MC4P_SIMPLETRANSFORMATION EXTENDS L_MC4P_TemplateTransformation
VAR
	SCSTORE : L_MC4P_IntermediateResultStore;
	SCSTORE_INTERNAL : L_MC4P_IntermediateResultStore;
END_VAR
END_FUNCTION_BLOCK

METHOD ADDTURNSTOJOINTS : L_IE1P_Error
VAR_INPUT
	PFLANGE_POS : POINTER TO ARRAY [1..6] OF LREAL;
	PJOINT_POS : POINTER TO ARRAY [1..6] OF LREAL;
END_VAR
VAR_IN_OUT
	SCTRAFOINFO : L_MC4P_TrafoInfo;
END_VAR
END_METHOD

METHOD CALCBACKWARDTRANSFORMATIONACC : L_IE1P_Error
VAR_INPUT
	PSTORE : POINTER TO L_MC4P_IntermediateResultStore;
END_VAR
VAR_IN_OUT
	SCTRAFOINFO : L_MC4P_TrafoInfo;
END_VAR
END_METHOD

METHOD CALCBACKWARDTRANSFORMATIONPOS : L_IE1P_Error
VAR_INPUT
	PSTORE : POINTER TO L_MC4P_IntermediateResultStore;
END_VAR
VAR_IN_OUT
	SCTRAFOINFO : L_MC4P_TrafoInfo;
END_VAR
END_METHOD

METHOD CALCBACKWARDTRANSFORMATIONVEL : L_IE1P_Error
VAR_INPUT
	PSTORE : POINTER TO L_MC4P_IntermediateResultStore;
END_VAR
VAR_IN_OUT
	SCTRAFOINFO : L_MC4P_TrafoInfo;
END_VAR
END_METHOD

METHOD CALCFORWARDTRANSFORMATIONACC : L_IE1P_Error
VAR_INPUT
	PSTORE : POINTER TO L_MC4P_IntermediateResultStore;
END_VAR
VAR_IN_OUT
	SCTRAFOINFO : L_MC4P_TrafoInfo;
END_VAR
END_METHOD

METHOD CALCFORWARDTRANSFORMATIONPOS : L_IE1P_Error
VAR_INPUT
	PSTORE : POINTER TO L_MC4P_IntermediateResultStore;
END_VAR
VAR_IN_OUT
	SCTRAFOINFO : L_MC4P_TrafoInfo;
END_VAR
END_METHOD

METHOD CALCFORWARDTRANSFORMATIONVEL : L_IE1P_Error
VAR_INPUT
	PSTORE : POINTER TO L_MC4P_IntermediateResultStore;
END_VAR
VAR_IN_OUT
	SCTRAFOINFO : L_MC4P_TrafoInfo;
END_VAR
END_METHOD

METHOD FB_INIT : BOOL
VAR_INPUT
	BINITRETAINS : BOOL;
	BINCOPYCODE : BOOL;
END_VAR
END_METHOD

METHOD CALCDINVERSEJACOBIAN : BOOL
VAR_INPUT
	ICOORDPROVIDER : L_MC4P_IKinCoordProvider;
	PDINVJACOBIAN : POINTER TO ARRAY [1..6, 1..6] OF LREAL;
END_VAR
VAR_OUTPUT
	SCERROR : L_MC4P_ErrorStruct;
END_VAR
END_METHOD

METHOD CALCDJACOBIAN : BOOL
VAR_INPUT
	ICOORDPROVIDER : L_MC4P_IKinCoordProvider;
	PDJACOBIAN : POINTER TO ARRAY [1..6, 1..6] OF LREAL;
END_VAR
VAR_OUTPUT
	SCERROR : L_MC4P_ErrorStruct;
END_VAR
END_METHOD

METHOD CALCINVERSEJACOBIAN : BOOL
VAR_INPUT
	ICOORDPROVIDER : L_MC4P_IKinCoordProvider;
	PINVJACOBIAN : POINTER TO ARRAY [1..6, 1..6] OF LREAL;
END_VAR
VAR_OUTPUT
	SCERROR : L_MC4P_ErrorStruct;
END_VAR
END_METHOD

METHOD CALCJACOBIAN : BOOL
VAR_INPUT
	ICOORDPROVIDER : L_MC4P_IKinCoordProvider;
	PJACOBIAN : POINTER TO ARRAY [1..6, 1..6] OF LREAL;
END_VAR
VAR_OUTPUT
	SCERROR : L_MC4P_ErrorStruct;
END_VAR
END_METHOD

METHOD MCS_ORIENTATIONCHECK : L_IE1P_Error
VAR_IN_OUT
	ICOORDPROVIDER : L_MC4P_KinCoordProvider;
END_VAR
END_METHOD

(* ---- L_MC4P_TCPFORCEOBSERVER.fb ---- *)
FUNCTION_BLOCK L_MC4P_TCPFORCEOBSERVER EXTENDS L_MC4P_Template_AG_KIN
VAR_INPUT
	XENABLE : BOOL;
	XUSEAXESGROUPPARAM : BOOL := FALSE;
	LRLOADMASS : LREAL;
	ITFDYNAMICPAR : L_MC4P_DynamicPar;
	LROBSERVATIONDYNAMIC : LREAL;
	EOBSERVATIONMODE : L_MC4P_ObservationMode;
END_VAR
VAR_OUTPUT
	XVALID : BOOL;
	XBUSY : BOOL;
	XERROR : BOOL;
	EERRORID : L_IE1P_Error;
	ALROBSERVEDTCPFORCE : ARRAY [1..3] OF LREAL;
	LROBSERVEDLOADMASS : LREAL;
END_VAR
VAR
	LICHANDLING : L_IMHP_LLMHandling;
	ALRGRAVITATION : ARRAY [1..3] OF LREAL;
	ALRCOULOMBFRIC : ARRAY [1..6] OF LREAL;
	ALRVISCFRIC : ARRAY [1..6] OF LREAL;
	ALRDYNAMICPAR : ARRAY [1..L_MC4P_Constants.uimaxNbrOfDynamicPar] OF LREAL;
	PLRREGRESSIONMATRIX : POINTER TO LREAL;
	XENABLEOLD : BOOL;
	EERRORTMP : L_IE1P_Error;
	ITFJACOBIAN : L_MC4P_IJacobi;
	ALRACTTORQUEACS : ARRAY [1..6] OF LREAL;
	ALRACTTORQUEJCS : ARRAY [1..6] OF LREAL;
	ALRCALCULATEDTORQUEJCS : ARRAY [1..6] OF LREAL;
	ALREXTTORQUE : ARRAY [1..6] OF LREAL;
	ALRTORQUEERROR : ARRAY [1..6] OF LREAL;
	ALRINVJACOBIAN : ARRAY [1..6, 1..6] OF LREAL;
	ALRTRANSPOSEDINVJACOBIAN : ARRAY [1..6, 1..6] OF LREAL;
	ALROBSERVEDTCPFORCEINT : ARRAY [1..6] OF LREAL;
	LROBSERVEDLOADMASSINT : LREAL;
	LROBSERVATIONDYNAMICLIM : LREAL;
	LROBSERVATIONDYNAMICINT : LREAL;
	APT1_ACTJCSPOS : ARRAY [1..6] OF L_USPP.L_USPP_PT1Filter;
	APT1_ACTJCSVEL : ARRAY [1..6] OF L_USPP.L_USPP_PT1Filter;
	APT1_ACTJCSACC : ARRAY [1..6] OF L_USPP.L_USPP_PT1Filter;
	APT1_ACTFCSPOS : ARRAY [1..6] OF L_USPP.L_USPP_PT1Filter;
	APT1_ACTFCSVEL : ARRAY [1..6] OF L_USPP.L_USPP_PT1Filter;
	APT1_ACTFCSACC : ARRAY [1..6] OF L_USPP.L_USPP_PT1Filter;
	APT1_ACTTORQUE : ARRAY [1..6] OF L_USPP.L_USPP_PT1Filter;
	AGOF : ARRAY [1..3] OF L_UMTP_GoodnessOfFit;
	LRCONVERGENCE : LREAL;
	LRVALIDTHRESHOLDON : LREAL := 0.75;
	LRVALIDTHRESHOLDOFF : LREAL := 0.5;
	RLS1 : L_UMTP_RLS;
	MASSMEANFILTER : L_MC4P_AvgValueFilter1D;
	AFORCEMEANFILTER : ARRAY [1..3] OF L_MC4P_AvgValueFilter1D;
	LRPT1FILTERTIME : LREAL;
	LRLAMBDA : LREAL;
	UIMEANFILTERTIME : UINT;
	XDIFFERENTIALDRIVE1ACTIVE : BOOL;
	PACTTRAFOEXTENSION1 : POINTER TO L_MC4P_TrafoExtensionBase;
	USINBROFDYNPAR : USINT;
	IDX : INT;
END_VAR
END_FUNCTION_BLOCK

METHOD CALCULATEMODEL
VAR_IN_OUT
	AXESGROUP : AXES_GROUP_KIN;
END_VAR
END_METHOD

(* ---- L_MC4P_TEACHCOORDINATESYSTEM.fb ---- *)
FUNCTION_BLOCK L_MC4P_TEACHCOORDINATESYSTEM EXTENDS L_MC4P_Template_AG_KIN
VAR_INPUT
	XEXECUTE : BOOL;
	XSTEPCONFIRM : BOOL;
	ECOORDSYSTEM : L_MC4P_CoordSystem;
END_VAR
VAR_OUTPUT
	XDONE : BOOL;
	XBUSY : BOOL;
	XERROR : BOOL;
	EERRORID : L_IE1P_Error;
	ENEXTSTEP : L_MC4P_TeachCoordinateSystemSteps;
	SCCOORDINATETRANSFORM : MC_COORD_REF;
END_VAR
VAR
	XEXECUTEOLD : BOOL;
	XSTEPCONFIRMOLD : BOOL;
	BASE_POS : ARRAY [1..3] OF LREAL;
	POS_TMP : ARRAY [1..3] OF LREAL;
	POS_TMP2 : ARRAY [1..3] OF LREAL;
	X_VEK : ARRAY [1..3] OF LREAL;
	Y_VEK : ARRAY [1..3] OF LREAL;
	Z_VEK : ARRAY [1..3] OF LREAL;
	XY_VEK : ARRAY [1..3] OF LREAL;
	T : ARRAY [1..4, 1..4] OF LREAL;
	MC_SETCOORDINATETRANSFORM1 : MC_SetCoordinateTransform;
END_VAR
END_FUNCTION_BLOCK

METHOD SETERROR
END_METHOD

(* ---- L_MC4P_TEMPLATE_AG_KIN.fb ---- *)
FUNCTION_BLOCK L_MC4P_TEMPLATE_AG_KIN EXTENDS L_MC4P_Template_ForAG
VAR_IN_OUT
	AXESGROUP : AXES_GROUP_KIN;
END_VAR
VAR
	SINSTANCESTR : STRING;
	AXESGROUP_WINITSTATEOLD : WORD;
END_VAR
END_FUNCTION_BLOCK

METHOD AXESGROUPINITDONE : BOOL
VAR_INPUT
	XEXECUTE : BOOL;
END_VAR
VAR_IN_OUT
	XERROR : BOOL;
	EERRORID : L_IE1P_Error;
	AXESGROUP : AXES_GROUP_KIN;
END_VAR
END_METHOD

METHOD FB_GETERRORITFID : DWORD
END_METHOD

METHOD FB_RESETERROR
VAR_INPUT
	XERROR : BOOL;
	WERRORID : WORD;
END_VAR
END_METHOD

METHOD FB_SETERROR
VAR_INPUT
	WERRORID : L_IE1P_Error := L_IE1P_Error.NoError;
	XSETERRORSTOP : BOOL := FALSE;
END_VAR
END_METHOD

METHOD FB_SETERRORINT
VAR_INPUT
	WERRORID : L_IE1P_Error := L_IE1P_Error.NoError;
	DWINTERNALID : DWORD;
	XSETERRORSTOP : BOOL := FALSE;
END_VAR
END_METHOD

METHOD FB_INIT : BOOL
VAR_INPUT
	BINITRETAINS : BOOL;
	BINCOPYCODE : BOOL;
END_VAR
END_METHOD

(* ---- L_MC4P_TEMPLATE_AG_KIN_LICENCE.fb ---- *)
FUNCTION_BLOCK L_MC4P_TEMPLATE_AG_KIN_LICENCE EXTENDS L_MC4P_Template_AG_KIN
VAR
	LICHANDLING : L_IMHP_LLMHandling;
	MC1P_LICENCE : L_MC1P_Template_Licence_150;
END_VAR
END_FUNCTION_BLOCK

METHOD ACTIVATEAPPCREDIT : BOOL
VAR_INPUT
	XACTIVATE : BOOL;
END_VAR
END_METHOD

(* ---- L_MC4P_TEMPLATE_AG_REF.fb ---- *)
FUNCTION_BLOCK L_MC4P_TEMPLATE_AG_REF EXTENDS L_MC4P_Template_ForAG
VAR_IN_OUT
	AXESGROUP : AXES_GROUP_REF;
END_VAR
VAR
	SINSTANCESTR : STRING;
	AXESGROUP_WINITSTATEOLD : WORD;
END_VAR
END_FUNCTION_BLOCK

METHOD AXESGROUPINITDONE : BOOL
VAR_INPUT
	XEXECUTE : BOOL;
END_VAR
VAR_IN_OUT
	XERROR : BOOL;
	EERRORID : L_IE1P_Error;
	AXESGROUP : AXES_GROUP_REF;
END_VAR
END_METHOD

METHOD FB_GETERRORITFID : DWORD
END_METHOD

METHOD FB_RESETERROR
VAR_INPUT
	XERROR : BOOL;
	WERRORID : WORD;
END_VAR
END_METHOD

METHOD FB_SETERROR
VAR_INPUT
	WERRORID : L_IE1P_Error := L_IE1P_Error.NoError;
	XSETERRORSTOP : BOOL := FALSE;
END_VAR
END_METHOD

METHOD FB_SETERRORINT
VAR_INPUT
	WERRORID : L_IE1P_Error := L_IE1P_Error.NoError;
	DWINTERNALID : DWORD;
	XSETERRORSTOP : BOOL := FALSE;
END_VAR
END_METHOD

METHOD FB_INIT : BOOL
VAR_INPUT
	BINITRETAINS : BOOL;
	BINCOPYCODE : BOOL;
END_VAR
END_METHOD

(* ---- L_MC4P_TEMPLATE_FORAG.fb ---- *)
FUNCTION_BLOCK L_MC4P_TEMPLATE_FORAG
VAR
	XERROROLD : BOOL;
	WERRORIDOLD : WORD;
	XDISABLEERRORRESET : BOOL;
	XDISABLEERRORLOGGING : BOOL;
	DWERRORITFID : DWORD;
	PFBBASEAXESGROUP : POINTER TO AXES_GROUP_REF;
	PSINSTANCESTR : POINTER TO STRING;
	DISABLEERRORLOGGING : BOOL;
	DISABLEERRORRESET : BOOL;
END_VAR
END_FUNCTION_BLOCK

METHOD SETINCTANCEINFO
VAR_INPUT
	PSINSTANCENAME : POINTER TO STRING;
	ERRORITFID : DWORD;
END_VAR
END_METHOD

METHOD SETINSTANCEINFOANDAXISPOINTER
VAR_INPUT
	PAXESGROUP : POINTER TO AXES_GROUP_REF;
	PSNAME : POINTER TO STRING;
END_VAR
END_METHOD

METHOD UPDATEAXISPOINTER
VAR_INPUT
	PAXESGROUP : POINTER TO AXES_GROUP_REF;
END_VAR
END_METHOD

METHOD FB_RESETERROR
VAR_INPUT
	XERROR : BOOL;
	WERRORID : WORD;
END_VAR
END_METHOD

METHOD FB_SETERROR
VAR_INPUT
	WERRORID : L_IE1P_Error := L_IE1P_Error.NoError;
	XSETERRORSTOP : BOOL := FALSE;
END_VAR
END_METHOD

METHOD FB_SETERRORINT
VAR_INPUT
	WERRORID : L_IE1P_Error := L_IE1P_Error.NoError;
	DWINTERNALID : DWORD;
	XSETERRORSTOP : BOOL := FALSE;
END_VAR
END_METHOD

(* ---- L_MC4P_TEMPLATE_KIN.fb ---- *)
FUNCTION_BLOCK L_MC4P_TEMPLATE_KIN
VAR
	SINSTANCESTR : STRING;
	XERROROLD : BOOL;
	WERRORIDOLD : WORD;
END_VAR
END_FUNCTION_BLOCK

METHOD FB_INIT : BOOL
VAR_INPUT
	BINITRETAINS : BOOL;
	BINCOPYCODE : BOOL;
END_VAR
END_METHOD

(* ---- L_MC4P_TEMPLATE_MOVE.fb ---- *)
FUNCTION_BLOCK L_MC4P_TEMPLATE_MOVE EXTENDS L_MC4P_Template_AG_KIN
VAR
	PMOVE : POINTER TO L_MC4P_MoveContPath;
	PROFILETIME : LREAL;
	REMAININGSEGMENTLENGTH : LREAL;
	REMAININGTIMEOFPROFILE : LREAL;
	TARGETREACHED : BOOL;
	TIMEIPOACTIVE : BOOL;
END_VAR
END_FUNCTION_BLOCK

METHOD GETREMAININGSEGMENTTIME : BOOL
VAR_INPUT
	LRDISTANCETOTARGET : LREAL;
END_VAR
VAR_OUTPUT
	LRREMAININGTIME : LREAL;
END_VAR
END_METHOD

METHOD FB_INIT : BOOL
VAR_INPUT
	BINITRETAINS : BOOL;
	BINCOPYCODE : BOOL;
END_VAR
END_METHOD

(* ---- L_MC4P_TEMPLATE_MOVE_FORSMARTFBS.fb ---- *)
FUNCTION_BLOCK L_MC4P_TEMPLATE_MOVE_FORSMARTFBS EXTENDS L_MC4P_Template_Move
VAR_IN_OUT
	FBMOVE : L_MC4P_MoveContPath;
END_VAR
VAR
	PMOVE : POINTER TO L_MC4P_MoveContPath;
END_VAR
END_FUNCTION_BLOCK

(* ---- L_MC4P_TEMPLATE_MOVELICENCE.fb ---- *)
FUNCTION_BLOCK L_MC4P_TEMPLATE_MOVELICENCE EXTENDS L_MC4P_Template_Move
VAR
	LICHANDLING : L_IMHP_LLMHandling;
	MC1P_LICENCE : L_MC1P_Template_Licence_150;
END_VAR
END_FUNCTION_BLOCK

METHOD ACTIVATEAPPCREDIT : BOOL
VAR_INPUT
	XACTIVATE : BOOL;
END_VAR
END_METHOD

(* ---- L_MC4P_TEMPLATETRANSFORMATION.fb ---- *)
FUNCTION_BLOCK L_MC4P_TEMPLATETRANSFORMATION
VAR_INPUT
	PAXESGROUP : POINTER TO AXES_GROUP_KIN;
END_VAR
VAR
	IDX : INT;
	ITRAFOEXTENSION1 : L_MC4P_ITrafoExtension;
	PTRAFOEXTENSION1 : POINTER TO L_MC4P_TrafoExtensionBase;
	PTOOLTRAFO : POINTER TO L_MC4P_ToolTrafo;
	PSTORE : POINTER TO L_MC4P_IntermediateResultStore;
	PSTORE_INTERNAL : POINTER TO L_MC4P_IntermediateResultStore;
	ALRACS2JCSSCALE : ARRAY [1..6] OF LREAL := [1.0, 1.0, 1.0, 1.0, 1.0, 1.0];
	ALRJCS2ACSSCALE : ARRAY [1..6] OF LREAL := [1.0, 1.0, 1.0, 1.0, 1.0, 1.0];
END_VAR
END_FUNCTION_BLOCK

METHOD COORD2ROBOTPOS
VAR_INPUT
	PCOORD : POINTER TO ARRAY [1..6] OF LREAL;
	ECONV : L_UMTP_RotationConvention;
	ROBOTPOS : REFERENCE TO L_UMTP_RobotPos;
	XISSI : BOOL;
END_VAR
END_METHOD

METHOD TOOLTRAFOFCSTOMCSACC
VAR_INPUT
	ICOORDPROVIDER : REFERENCE TO L_MC4P_KinCoordProvider;
	BVALIDFRAME : BOOL;
	ETOOLSYSTEM : L_MC4P_ToolSystem;
END_VAR
END_METHOD

METHOD TOOLTRAFOFCSTOMCSPOS : L_MC4P_ErrorStruct
VAR_INPUT
	ICOORDPROVIDER : REFERENCE TO L_MC4P_KinCoordProvider;
	BVALIDFRAME : BOOL;
	ETOOLSYSTEM : L_MC4P_ToolSystem;
END_VAR
END_METHOD

METHOD TOOLTRAFOFCSTOMCSVEL
VAR_INPUT
	ICOORDPROVIDER : REFERENCE TO L_MC4P_KinCoordProvider;
	BVALIDFRAME : BOOL;
	ETOOLSYSTEM : L_MC4P_ToolSystem;
END_VAR
END_METHOD

METHOD TOOLTRAFOMCSTOFCSACC
VAR_INPUT
	ICOORDPROVIDER : REFERENCE TO L_MC4P_KinCoordProvider;
	BVALIDFRAME : BOOL;
	ETOOLSYSTEM : L_MC4P_ToolSystem;
END_VAR
END_METHOD

METHOD TOOLTRAFOMCSTOFCSPOS : L_MC4P_ErrorStruct
VAR_INPUT
	ICOORDPROVIDER : REFERENCE TO L_MC4P_KinCoordProvider;
	BVALIDFRAME : BOOL;
	ETOOLSYSTEM : L_MC4P_ToolSystem;
END_VAR
END_METHOD

METHOD TOOLTRAFOMCSTOFCSVEL
VAR_INPUT
	ICOORDPROVIDER : REFERENCE TO L_MC4P_KinCoordProvider;
	BVALIDFRAME : BOOL;
	ETOOLSYSTEM : L_MC4P_ToolSystem;
END_VAR
END_METHOD

METHOD TRAFOMCSTOWCSACC
VAR_INPUT
	ICOORDPROVIDER : REFERENCE TO L_MC4P_KinCoordProvider;
	BVALIDFRAME : BOOL;
END_VAR
END_METHOD

METHOD TRAFOMCSTOWCSPOS : L_MC4P_ErrorStruct
VAR_INPUT
	ICOORDPROVIDER : REFERENCE TO L_MC4P_KinCoordProvider;
	BVALIDFRAME : BOOL;
END_VAR
END_METHOD

METHOD TRAFOMCSTOWCSVEL
VAR_INPUT
	ICOORDPROVIDER : REFERENCE TO L_MC4P_KinCoordProvider;
	BVALIDFRAME : BOOL;
END_VAR
END_METHOD

METHOD TRAFOWCSTOMCSACC
VAR_INPUT
	ICOORDPROVIDER : REFERENCE TO L_MC4P_KinCoordProvider;
	BVALIDFRAME : BOOL;
END_VAR
END_METHOD

METHOD TRAFOWCSTOMCSPOS : L_MC4P_ErrorStruct
VAR_INPUT
	ICOORDPROVIDER : REFERENCE TO L_MC4P_KinCoordProvider;
	BVALIDFRAME : BOOL;
END_VAR
END_METHOD

METHOD TRAFOWCSTOMCSVEL
VAR_INPUT
	ICOORDPROVIDER : REFERENCE TO L_MC4P_KinCoordProvider;
	BVALIDFRAME : BOOL;
END_VAR
END_METHOD

METHOD CALCDINVERSEJACOBIAN : BOOL
VAR_INPUT
	ICOORDPROVIDER : L_MC4P_IKinCoordProvider;
	PDINVJACOBIAN : POINTER TO ARRAY [1..6, 1..6] OF LREAL;
END_VAR
VAR_OUTPUT
	SCERROR : L_MC4P_ErrorStruct;
END_VAR
END_METHOD

METHOD CALCDJACOBIAN : BOOL
VAR_INPUT
	ICOORDPROVIDER : L_MC4P_IKinCoordProvider;
	PDJACOBIAN : POINTER TO ARRAY [1..6, 1..6] OF LREAL;
END_VAR
VAR_OUTPUT
	SCERROR : L_MC4P_ErrorStruct;
END_VAR
END_METHOD

METHOD CALCINVERSEJACOBIAN : BOOL
VAR_INPUT
	ICOORDPROVIDER : L_MC4P_IKinCoordProvider;
	PINVJACOBIAN : POINTER TO ARRAY [1..6, 1..6] OF LREAL;
END_VAR
VAR_OUTPUT
	SCERROR : L_MC4P_ErrorStruct;
END_VAR
END_METHOD

METHOD CALCJACOBIAN : BOOL
VAR_INPUT
	ICOORDPROVIDER : L_MC4P_IKinCoordProvider;
	PJACOBIAN : POINTER TO ARRAY [1..6, 1..6] OF LREAL;
END_VAR
VAR_OUTPUT
	SCERROR : L_MC4P_ErrorStruct;
END_VAR
END_METHOD

METHOD CALCNUMERICALINVERSEJACOBIAN : L_IE1P_Error
VAR_INPUT
	ICOORDPROVIDER : L_MC4P_IKinCoordProvider;
	PINVJACOBIAN : POINTER TO ARRAY [1..6, 1..6] OF LREAL;
END_VAR
END_METHOD

METHOD CALCNUMERICALJACOBIAN : L_IE1P_Error
VAR_INPUT
	ICOORDPROVIDER : L_MC4P_IKinCoordProvider;
	PJACOBIAN : POINTER TO ARRAY [1..6, 1..6] OF LREAL;
END_VAR
END_METHOD

METHOD BWDACC : BOOL
VAR_INPUT
	ICOORDPROVIDER : REFERENCE TO L_MC4P_KinCoordProvider;
END_VAR
VAR_OUTPUT
	SCERROR : L_MC4P_ErrorStruct;
END_VAR
VAR_IN_OUT
	SCTRAFOINFO : L_MC4P_TrafoInfo;
END_VAR
END_METHOD

METHOD BWDPOS : BOOL
VAR_INPUT
	ICOORDPROVIDER : REFERENCE TO L_MC4P_KinCoordProvider;
END_VAR
VAR_OUTPUT
	SCERROR : L_MC4P_ErrorStruct;
END_VAR
VAR_IN_OUT
	SCTRAFOINFO : L_MC4P_TrafoInfo;
END_VAR
END_METHOD

METHOD BWDVEL : BOOL
VAR_INPUT
	ICOORDPROVIDER : REFERENCE TO L_MC4P_KinCoordProvider;
END_VAR
VAR_OUTPUT
	SCERROR : L_MC4P_ErrorStruct;
END_VAR
VAR_IN_OUT
	SCTRAFOINFO : L_MC4P_TrafoInfo;
END_VAR
END_METHOD

METHOD CALCPASSIVEJOINTS : L_IE1P_Error
VAR_INPUT
	PFLANGE_POS : POINTER TO ARRAY [1..6] OF LREAL;
	PJOINT_POS : POINTER TO ARRAY [1..6] OF LREAL;
	PPASSIVEJOINT_POS : POINTER TO ARRAY [1..6, 1..3] OF LREAL;
END_VAR
END_METHOD

METHOD CALCULATECONFIGURATION : L_IE1P_Error
VAR_INPUT
	PJOINT_POS : POINTER TO ARRAY [1..6] OF LREAL;
END_VAR
VAR_IN_OUT
	SCTRAFOINFO : L_MC4P_TrafoInfo;
END_VAR
END_METHOD

METHOD FWDACC : BOOL
VAR_INPUT
	ICOORDPROVIDER : REFERENCE TO L_MC4P_KinCoordProvider;
END_VAR
VAR_OUTPUT
	SCERROR : L_MC4P_ErrorStruct;
END_VAR
VAR_IN_OUT
	SCTRAFOINFO : L_MC4P_TrafoInfo;
END_VAR
END_METHOD

METHOD FWDPOS : BOOL
VAR_INPUT
	ICOORDPROVIDER : REFERENCE TO L_MC4P_KinCoordProvider;
END_VAR
VAR_OUTPUT
	SCERROR : L_MC4P_ErrorStruct;
END_VAR
VAR_IN_OUT
	SCTRAFOINFO : L_MC4P_TrafoInfo;
END_VAR
END_METHOD

METHOD FWDVEL : BOOL
VAR_INPUT
	ICOORDPROVIDER : REFERENCE TO L_MC4P_KinCoordProvider;
END_VAR
VAR_OUTPUT
	SCERROR : L_MC4P_ErrorStruct;
END_VAR
VAR_IN_OUT
	SCTRAFOINFO : L_MC4P_TrafoInfo;
END_VAR
END_METHOD

METHOD GETTRAFOEXTENSION1 : L_MC4P_ITrafoExtension
VAR_OUTPUT
	PFB : POINTER TO L_MC4P_TrafoExtensionBase;
END_VAR
END_METHOD

METHOD MCS_ORIENTATIONCHECK : L_IE1P_Error
VAR_IN_OUT
	ICOORDPROVIDER : L_MC4P_KinCoordProvider;
END_VAR
END_METHOD

METHOD SETTRAFOEXTENSION1
VAR_INPUT
	TRAFOEXTENSION : L_MC4P_ITrafoExtension;
	PFB : POINTER TO L_MC4P_TrafoExtensionBase;
END_VAR
END_METHOD

METHOD CHECKNEIGHBOURHOOD : L_IE1P_Error
VAR_INPUT
	PJOINT_POS : POINTER TO ARRAY [1..6] OF LREAL;
END_VAR
VAR_IN_OUT
	SCTRAFOINFO : L_MC4P_TrafoInfo;
END_VAR
END_METHOD

METHOD COUNTREVOLUTIONSFORWARDTRAFO : L_IE1P_Error
VAR_INPUT
	PJOINT_POS : POINTER TO ARRAY [1..6] OF LREAL;
END_VAR
VAR_IN_OUT
	SCTRAFOINFO : L_MC4P_TrafoInfo;
END_VAR
END_METHOD

METHOD IDENTIFYTRAFOCASE : L_IE1P_Error
VAR_INPUT
	PKART_POS : POINTER TO ARRAY [1..6] OF LREAL;
	PMCS_POS : POINTER TO ARRAY [1..6] OF LREAL;
	PFLANGE_POS : POINTER TO ARRAY [1..6] OF LREAL;
	PJOINT_POS : POINTER TO ARRAY [1..6] OF LREAL;
	PAXES_POS : POINTER TO ARRAY [1..6] OF LREAL;
END_VAR
VAR_IN_OUT
	ILOWERSYSTEM : INT;
	IUPPERSYSTEM : INT;
END_VAR
END_METHOD

METHOD PRELOADCONSTANTAXES
VAR_INPUT
	PACSPOS : POINTER TO ARRAY [1..6] OF LREAL;
	PJCSPOS : POINTER TO ARRAY [1..6] OF LREAL;
	PFCSPOS : POINTER TO ARRAY [1..6] OF LREAL;
	PMCSPOS : POINTER TO ARRAY [1..6] OF LREAL;
	PWCSPOS : POINTER TO ARRAY [1..6] OF LREAL;
END_VAR
VAR_IN_OUT
	SCTRAFOINFO : L_MC4P_TrafoInfo;
END_VAR
END_METHOD

METHOD ADDTURNSTOJOINTS : L_IE1P_Error
VAR_INPUT
	PFLANGE_POS : POINTER TO ARRAY [1..6] OF LREAL;
	PJOINT_POS : POINTER TO ARRAY [1..6] OF LREAL;
END_VAR
VAR_IN_OUT
	SCTRAFOINFO : L_MC4P_TrafoInfo;
END_VAR
END_METHOD

METHOD CALCBACKWARDTRANSFORMATIONACC : L_IE1P_Error
VAR_INPUT
	PSTORE : POINTER TO L_MC4P_IntermediateResultStore;
END_VAR
VAR_IN_OUT
	SCTRAFOINFO : L_MC4P_TrafoInfo;
END_VAR
END_METHOD

METHOD CALCBACKWARDTRANSFORMATIONPOS : L_IE1P_Error
VAR_INPUT
	PSTORE : POINTER TO L_MC4P_IntermediateResultStore;
END_VAR
VAR_IN_OUT
	SCTRAFOINFO : L_MC4P_TrafoInfo;
END_VAR
END_METHOD

METHOD CALCBACKWARDTRANSFORMATIONVEL : L_IE1P_Error
VAR_INPUT
	PSTORE : POINTER TO L_MC4P_IntermediateResultStore;
END_VAR
VAR_IN_OUT
	SCTRAFOINFO : L_MC4P_TrafoInfo;
END_VAR
END_METHOD

METHOD CALCFORWARDTRANSFORMATIONACC : L_IE1P_Error
VAR_INPUT
	PSTORE : POINTER TO L_MC4P_IntermediateResultStore;
END_VAR
VAR_IN_OUT
	SCTRAFOINFO : L_MC4P_TrafoInfo;
END_VAR
END_METHOD

METHOD CALCFORWARDTRANSFORMATIONPOS : L_IE1P_Error
VAR_INPUT
	PSTORE : POINTER TO L_MC4P_IntermediateResultStore;
END_VAR
VAR_IN_OUT
	SCTRAFOINFO : L_MC4P_TrafoInfo;
END_VAR
END_METHOD

METHOD CALCFORWARDTRANSFORMATIONVEL : L_IE1P_Error
VAR_INPUT
	PSTORE : POINTER TO L_MC4P_IntermediateResultStore;
END_VAR
VAR_IN_OUT
	SCTRAFOINFO : L_MC4P_TrafoInfo;
END_VAR
END_METHOD

METHOD CALCPASSIVEJOINTSACC : L_IE1P_Error
VAR_INPUT
	PSTORE : POINTER TO L_MC4P_IntermediateResultStore;
END_VAR
VAR_IN_OUT
	SCTRAFOINFO : L_MC4P_TrafoInfo;
END_VAR
END_METHOD

METHOD CALCPASSIVEJOINTSPOS : L_IE1P_Error
VAR_INPUT
	PSTORE : POINTER TO L_MC4P_IntermediateResultStore;
END_VAR
VAR_IN_OUT
	SCTRAFOINFO : L_MC4P_TrafoInfo;
END_VAR
END_METHOD

METHOD CALCPASSIVEJOINTSVEL : L_IE1P_Error
VAR_INPUT
	PSTORE : POINTER TO L_MC4P_IntermediateResultStore;
END_VAR
VAR_IN_OUT
	SCTRAFOINFO : L_MC4P_TrafoInfo;
END_VAR
END_METHOD

METHOD FINALIZEBWD : L_IE1P_Error
VAR_IN_OUT
	SCTRAFOINFO : L_MC4P_TrafoInfo;
	ICOORDPROVIDER : L_MC4P_KinCoordProvider;
END_VAR
END_METHOD

METHOD TRANSFORMREVOLUTEJOINTS : L_IE1P_Error
VAR_INPUT
	PJCSPOS : POINTER TO ARRAY [1..6] OF LREAL;
END_VAR
VAR_IN_OUT
	SCTRAFOINFO : L_MC4P_TrafoInfo;
END_VAR
END_METHOD

(* ---- L_MC4P_TOOLCONTROL.fb ---- *)
FUNCTION_BLOCK L_MC4P_TOOLCONTROL
VAR_INPUT
	XENABLE : BOOL;
	ETOOLSYSTEM : L_MC4P_ToolSystem;
END_VAR
VAR_OUTPUT
	XBUSY : BOOL;
	XERROR : BOOL;
	EERRORID : L_IE1P_Error;
	XPULSEON : BOOL;
	XPULSEOFF : BOOL;
	LRTIMETOPULSE : LREAL;
END_VAR
VAR_IN_OUT
	AXESGROUP : AXES_GROUP_KIN;
END_VAR
VAR
	_ON_TRIG : R_Trig;
	_OFF_TRIG : R_Trig;
	_ITFTOOL : L_MC4P_IToolInfo;
	_NSTATE : DWORD := 10;
	_ETOOLSYSTEMFREEZE : L_MC4P_ToolSystem;
	_PTOOL : POINTER TO L_MC4P_ToolTrafo;
	_ETOOLREQU : L_MC4P_ToolRequest;
	_LRSWITCHTIME : LREAL;
	_MODEL : L_UBUP_BehaviourModel_LCon;
END_VAR
END_FUNCTION_BLOCK

METHOD CYCLICACTION
VAR_INPUT
	ITFTIMINGCONTROLLER : L_UBUP.L_UBUP_ITimingController;
END_VAR
VAR_OUTPUT
	XCOMPLETE : BOOL;
	XABORT : BOOL;
	IERRORID : INT;
END_VAR
END_METHOD

METHOD FINALIZEACTION
VAR_INPUT
	XABORTPROPOSED : BOOL;
	IERRORIDPROPOSED : INT;
END_VAR
VAR_OUTPUT
	XCOMPLETE : BOOL;
	XABORT : BOOL;
	IERRORID : INT;
END_VAR
END_METHOD

METHOD RESETACTION
VAR_OUTPUT
	XCOMPLETE : BOOL;
END_VAR
END_METHOD

METHOD STARTACTION
VAR_OUTPUT
	XCOMPLETE : BOOL;
	IERRORID : INT;
END_VAR
END_METHOD

(* ---- L_MC4P_TOOLTRAFO.fb ---- *)
FUNCTION_BLOCK L_MC4P_TOOLTRAFO
VAR_INPUT
	TOOLPARAM : L_MC4P_TOOL_REF;
	EROTATIONCONVENTION : L_UMTP_RotationConvention;
	ISWITCHONTIME : INT;
	ISWITCHOFFTIME : INT;
END_VAR
VAR_OUTPUT
	T_01 : ARRAY [1..4, 1..4] OF LREAL;
	T_01_FRAME : L_UMTP_RobotFrame;
	T_10 : ARRAY [1..4, 1..4] OF LREAL;
	T_10_FRAME : L_UMTP_RobotFrame;
END_VAR
VAR
	TOOLPARAMINT : L_MC4P_TOOL_REF;
	EROTATIONCONVENTIONINT : L_UMTP_RotationConvention;
	PAXESGROUP : POINTER TO AXES_GROUP_KIN;
END_VAR
END_FUNCTION_BLOCK

METHOD CALCHOMTRAFO
VAR_IN_OUT
	AXESGROUP : AXES_GROUP_KIN;
END_VAR
END_METHOD

METHOD ROTATE_FCS2TCS
VAR_INPUT
	PALRIN : POINTER TO ARRAY [1..6] OF LREAL;
	PALROUT : POINTER TO ARRAY [1..6] OF LREAL;
END_VAR
END_METHOD

METHOD ROTATE_TCS2FCS
VAR_INPUT
	PALRIN : POINTER TO ARRAY [1..6] OF LREAL;
	PALROUT : POINTER TO ARRAY [1..6] OF LREAL;
END_VAR
END_METHOD

(* ---- L_MC4P_TRACELIST.fb ---- *)
FUNCTION_BLOCK L_MC4P_TRACELIST
VAR_INPUT
	XENABLE : BOOL;
	PAXESGROUP : POINTER TO AXES_GROUP_KIN;
END_VAR
VAR
	PLISTELEMENT : POINTER TO L_MC4P_ListElement;
	VISULISTTABLE : ARRAY [0..L_MC4P_Constants.SizeVisuArray] OF L_MC4P_VisuListTableData;
	BFINISHED : BOOL := 0;
	IINDEX : INT := 0;
	XREADFROMLISTELEMENTLAST : BOOL := TRUE;
	HEVENTCOMMCYCLE : Systypes.RTS_IEC_HANDLE := SysTypes.RTS_INVALID_HANDLE;
	HINTERFACECOMMCYCLE : Systypes.RTS_IEC_HANDLE := SysTypes.RTS_INVALID_HANDLE;
	ITFCALLBACK : CmpEventMgr.ICmpEventCallback;
	DWEVENTCOUNTER : DWORD;
END_VAR
END_FUNCTION_BLOCK

METHOD FILLVISULISTTABLEELEMENT
END_METHOD

METHOD MAIN
END_METHOD

METHOD EVENTCALLBACK : UDINT
VAR_INPUT
	PEVENTPARAM : POINTER TO EventParam;
END_VAR
END_METHOD

METHOD REGISTEREVENT
END_METHOD

METHOD UNREGISTEREVENT
END_METHOD

(* ---- L_MC4P_TRACKCONVEYORBELT_INTERNAL.fb ---- *)
FUNCTION_BLOCK L_MC4P_TRACKCONVEYORBELT_INTERNAL EXTENDS L_MC4P_TrackKinematics
VAR_INPUT
	ITFCONVEYORBELT : L_MC1P_IAXIS_REF_MASTERVALUES;
	EXECUTE : BOOL;
	ABORT : BOOL;
	CONVEYORBELTORIGIN : ARRAY [1..6] OF LREAL;
	INITIALOBJECTPOSITION : ARRAY [1..6] OF LREAL;
	COORDSYSTEM : L_MC4P_CoordSystem;
	COORDTYPE : L_MC4P_CoordType;
	CLUTCHDISTANCE : LREAL;
	CLUTCHTIME : LREAL;
	CLUTCHTIMEABORT : LREAL;
	SETDYNPCS : BOOL := TRUE;
END_VAR
VAR_OUTPUT
	DONE : BOOL;
	BUSY : BOOL;
	ACTIVE : BOOL;
	COMMANDABORTED : BOOL;
	ERROR : BOOL;
	ERRORID : L_IE1P_Error;
	INSYNC : BOOL;
	DYNAMICPCSSET : BOOL;
END_VAR
VAR
	LRCONVBELTPOSITIONOLD : LREAL := 0;
	LRCOUNTEDMODULOCYCLES : LREAL := 0;
	EMASTERDIRECTIONSAVED : MC_Direction := MC_Direction.mcPositiveDirection;
	XMASTERVALID : BOOL;
	FBCONSIDERCVUNSTEADY : L_MC1P_ConsiderMasterUnsteady;
	CLUTCHEXTERNAL : LREAL;
END_VAR
END_FUNCTION_BLOCK

METHOD GETCLUTCHPARAMETER : BOOL
VAR_OUTPUT
	EERRORID : L_IE1P_Error;
END_VAR
END_METHOD

METHOD GETINITOBJPOS : MC_Coord_Ref
END_METHOD

METHOD GETMASTERDIRECTION : BOOL
VAR_INPUT
	ITFCONVEYORBELT : L_MC1P_IAXIS_REF_MASTERVALUES;
END_VAR
END_METHOD

METHOD GETMASTERVALUES : BOOL
VAR_INPUT
	PALRINITMASTERPOS : POINTER TO ARRAY [1..6] OF LREAL;
	PASCCNVVALUESCCS : POINTER TO ARRAY [1..6] OF L_MC4P_AxisProfile;
	PASCCNVVALUESCCSOLD : POINTER TO ARRAY [1..6] OF L_MC4P_AxisProfile;
	LRMASTERPOSEXTRAPOL : LREAL;
END_VAR
END_METHOD

METHOD MAIN
VAR_INPUT
	ITFCONVEYORBELT : L_MC1P_IAXIS_REF_MASTERVALUES;
END_VAR
VAR_IN_OUT
	AXESGROUP : AXES_GROUP_KIN;
	FBBASE : L_MC4P_Template_AG_KIN;
END_VAR
END_METHOD

METHOD PARAMETERFREEZE
VAR_OUTPUT
	EERRORID : L_IE1P_Error;
END_VAR
VAR_IN_OUT
	AXESGROUP : AXES_GROUP_KIN;
	FBBASE : L_MC4P_Template_AG_KIN;
END_VAR
END_METHOD

METHOD SYNCINONPOS : BOOL
VAR_INPUT
	PASCCNVVALUESCCS : POINTER TO ARRAY [1..6] OF L_MC4P_AxisProfile;
	ALRSUPERPOSPOSATCLUTCH : ARRAY [1..3] OF LREAL;
	PTRAFO_BASE_MCS : POINTER TO L_MC4P_CoordTrafo;
	LRCLUTCHDISTANCE : LREAL;
END_VAR
VAR_OUTPUT
	XINSYNC : BOOL;
END_VAR
VAR_IN_OUT
	AXESGROUP : AXES_GROUP_KIN;
	FBBASE : L_MC4P_Template_AG_KIN;
END_VAR
END_METHOD

METHOD SYNCINONTIME : BOOL
VAR_INPUT
	PASCCNVVALUESCCS : POINTER TO ARRAY [1..6] OF L_MC4P_AxisProfile;
	ALRSUPERPOSPOSATCLUTCH : ARRAY [1..3] OF LREAL;
	PTRAFO_BASE_MCS : POINTER TO L_MC4P_CoordTrafo;
	LRCLUTCHDISTANCE : LREAL;
END_VAR
VAR_OUTPUT
	XINSYNC : BOOL;
END_VAR
VAR_IN_OUT
	AXESGROUP : AXES_GROUP_KIN;
	FBBASE : L_MC4P_Template_AG_KIN;
END_VAR
END_METHOD

METHOD SYNCOUTONPOS : BOOL
VAR_INPUT
	PASCCNVVALUESCCS : POINTER TO ARRAY [1..6] OF L_MC4P_AxisProfile;
	ALRSUPERPOSPOSATCLUTCH : ARRAY [1..3] OF LREAL;
	PTRAFO_BASE_MCS : POINTER TO L_MC4P_CoordTrafo;
	LRCLUTCHDISTANCE : LREAL;
END_VAR
VAR_OUTPUT
	XSYNCOUTDONE : BOOL;
END_VAR
VAR_IN_OUT
	AXESGROUP : AXES_GROUP_KIN;
	FBBASE : L_MC4P_Template_AG_KIN;
END_VAR
END_METHOD

METHOD SYNCOUTONTIME : BOOL
VAR_INPUT
	PASCCNVVALUESCCS : POINTER TO ARRAY [1..6] OF L_MC4P_AxisProfile;
	ALRSUPERPOSPOSATCLUTCH : ARRAY [1..3] OF LREAL;
	PTRAFO_BASE_MCS : POINTER TO L_MC4P_CoordTrafo;
	LRCLUTCHDISTANCE : LREAL;
	XSYNCOUTKEEPPOSITION : BOOL;
END_VAR
VAR_OUTPUT
	XSYNCOUTDONE : BOOL;
END_VAR
VAR_IN_OUT
	AXESGROUP : AXES_GROUP_KIN;
	FBBASE : L_MC4P_Template_AG_KIN;
END_VAR
END_METHOD

METHOD SYNCHRON : BOOL
VAR_INPUT
	PASCCNVVALUESCCS : POINTER TO ARRAY [1..6] OF L_MC4P_AxisProfile;
	PTRAFO_BASE_MCS : POINTER TO L_MC4P_CoordTrafo;
END_VAR
END_METHOD

(* ---- L_MC4P_TRACKKINEMATICS.fb ---- *)
FUNCTION_BLOCK L_MC4P_TRACKKINEMATICS
VAR_INPUT
	EMASTERVALUESOURCE : MC_SOURCE := MC_SOURCE.mcCommandedValue;
END_VAR
VAR
	XDONE_INTERN : BOOL;
	XBUSY_INTERN : BOOL;
	XACTIVE_INTERN : BOOL;
	XCOMMANDABORTED_INTERN : BOOL;
	XERROR_INTERN : BOOL;
	EERRORID_INTERN : L_IE1P_Error;
	XINSYNC_INTERN : BOOL;
	DYNAMICPCSSET_INTERN : BOOL;
	WSTEP : L_MC4P_TrackKinematicsStates;
	WSTEPOLD : L_MC4P_TrackKinematicsStates;
	XEXECUTEOLD : BOOL;
	XSETDYNPCSINDEPENDANTOLD : BOOL;
	XCALCDYNPCS : BOOL;
	XERRORLASTCYCLE : BOOL;
	XABORTOLD : BOOL;
	XABORTEDMOVEMENT : BOOL;
	XABORTFB : BOOL;
	XRESTARTSYNC : BOOL;
	XWINSTANCE : __XWORD;
	SCINPUTPARAM : L_MC4P_TrackInputParam;
	PSCSUPERPOSDATA : POINTER TO L_MC4P_SuperposHandler;
	SCINITIALPCSINTERN : L_MC4P_CoordTrafo;
	PSCHANDSHAKE : POINTER TO L_MC4P_TrackingHandshake;
	ASCCONVEYORVALUES : ARRAY [1..6] OF L_MC4P_AxisProfile;
	ASCCONVEYORVALUESFIXED : ARRAY [1..6] OF L_MC4P_AxisProfile;
	ASCCONVEYORVALUESOLD : ARRAY [1..6] OF L_MC4P_AxisProfile;
	XCLUTCHINITDONE : BOOL;
	ASCENDSLAVE : ARRAY [1..7] OF L_MC4P_AxisProfile;
	ASCSTARTSLAVE : ARRAY [1..7] OF L_MC4P_AxisProfile;
	ALRMASTERCLUTCHPOS : ARRAY [1..6] OF LREAL;
	ACLUTCHFB : ARRAY [1..7] OF L_MC4P_Clutch;
	ALRCNVPOSATCLINCCS : ARRAY [1..6] OF LREAL;
	ALRSUPERPOSPOSTEMP : ARRAY [1..3] OF LREAL;
	LRTIMECOUNTER : LREAL;
	LRCLUTCHTIMEABORTDEFAULT : LREAL := 1.0;
	LRCLUTCHEXTERNAL : LREAL := -1.0;
	XUSECLUTCHEXTERNAL : BOOL;
	ASCSLAVEEXTRAPOL : ARRAY [1..7] OF L_MC4P_AxisProfile;
	ALRACCMINUS0 : ARRAY [1..7] OF LREAL;
	ALRVELMINUS0 : ARRAY [1..7] OF LREAL;
	ALRVELMINUS1 : ARRAY [1..7] OF LREAL;
	ALRPOSMINUS0 : ARRAY [1..7] OF LREAL;
	ALRPOSMINUS1 : ARRAY [1..7] OF LREAL;
	ALRPOSMINUS2 : ARRAY [1..7] OF LREAL;
	XABORTAGSTOPPING : BOOL;
	XSTATEMACHINE : BOOL;
	MASTERVALUESOURCE : MC_SOURCE;
END_VAR
END_FUNCTION_BLOCK

METHOD CALCDYNPCS : BOOL
VAR_INPUT
	BINITIALCALL : BOOL;
	PASCACTCNVVALUESCCS : POINTER TO ARRAY [1..6] OF L_MC4P_AxisProfile;
END_VAR
VAR_IN_OUT
	AXESGROUP : AXES_GROUP_KIN;
	FBBASE : L_MC4P_Template_AG_KIN;
END_VAR
END_METHOD

METHOD FB_INIT : BOOL
VAR_INPUT
	BINITRETAINS : BOOL;
	BINCOPYCODE : BOOL;
END_VAR
END_METHOD

METHOD GETCLUTCHPARAMETER : BOOL
VAR_OUTPUT
	EERRORID : L_IE1P_Error;
END_VAR
END_METHOD

METHOD GETINITOBJPOS : MC_Coord_Ref
END_METHOD

METHOD GETMASTERVALUES : BOOL
VAR_INPUT
	PALRINITMASTERPOS : POINTER TO ARRAY [1..6] OF LREAL;
	PASCCNVVALUESCCS : POINTER TO ARRAY [1..6] OF L_MC4P_AxisProfile;
	PASCCNVVALUESCCSOLD : POINTER TO ARRAY [1..6] OF L_MC4P_AxisProfile;
	LRMASTERPOSEXTRAPOL : LREAL;
END_VAR
END_METHOD

METHOD PARAMETERFREEZE
VAR_OUTPUT
	EERRORID : L_IE1P_Error;
END_VAR
VAR_IN_OUT
	AXESGROUP : AXES_GROUP_KIN;
	FBBASE : L_MC4P_Template_AG_KIN;
END_VAR
END_METHOD

METHOD PASSTHROUGHTRACKINGOFFSETRESET : BOOL
VAR_IN_OUT
	AXESGROUP : AXES_GROUP_KIN;
	FBBASE : L_MC4P_Template_AG_KIN;
END_VAR
END_METHOD

METHOD RESETSUPERPOSCLUTCHINITDONE
END_METHOD

METHOD SETCONVEYORVALUESFIXED
END_METHOD

METHOD SYNCINONPOS : BOOL
VAR_INPUT
	PASCCNVVALUESCCS : POINTER TO ARRAY [1..6] OF L_MC4P_AxisProfile;
	ALRSUPERPOSPOSATCLUTCH : ARRAY [1..3] OF LREAL;
	PTRAFO_BASE_MCS : POINTER TO L_MC4P_CoordTrafo;
	LRCLUTCHDISTANCE : LREAL;
END_VAR
VAR_OUTPUT
	XINSYNC : BOOL;
END_VAR
VAR_IN_OUT
	AXESGROUP : AXES_GROUP_KIN;
	FBBASE : L_MC4P_Template_AG_KIN;
END_VAR
END_METHOD

METHOD SYNCINONTIME : BOOL
VAR_INPUT
	PASCCNVVALUESCCS : POINTER TO ARRAY [1..6] OF L_MC4P_AxisProfile;
	ALRSUPERPOSPOSATCLUTCH : ARRAY [1..3] OF LREAL;
	PTRAFO_BASE_MCS : POINTER TO L_MC4P_CoordTrafo;
	LRCLUTCHDISTANCE : LREAL;
END_VAR
VAR_OUTPUT
	XINSYNC : BOOL;
END_VAR
VAR_IN_OUT
	AXESGROUP : AXES_GROUP_KIN;
	FBBASE : L_MC4P_Template_AG_KIN;
END_VAR
END_METHOD

METHOD SYNCOUTONPOS : BOOL
VAR_INPUT
	PASCCNVVALUESCCS : POINTER TO ARRAY [1..6] OF L_MC4P_AxisProfile;
	ALRSUPERPOSPOSATCLUTCH : ARRAY [1..3] OF LREAL;
	PTRAFO_BASE_MCS : POINTER TO L_MC4P_CoordTrafo;
	LRCLUTCHDISTANCE : LREAL;
END_VAR
VAR_OUTPUT
	XSYNCOUTDONE : BOOL;
END_VAR
VAR_IN_OUT
	AXESGROUP : AXES_GROUP_KIN;
	FBBASE : L_MC4P_Template_AG_KIN;
END_VAR
END_METHOD

METHOD SYNCOUTONTIME : BOOL
VAR_INPUT
	PASCCNVVALUESCCS : POINTER TO ARRAY [1..6] OF L_MC4P_AxisProfile;
	ALRSUPERPOSPOSATCLUTCH : ARRAY [1..3] OF LREAL;
	PTRAFO_BASE_MCS : POINTER TO L_MC4P_CoordTrafo;
	LRCLUTCHDISTANCE : LREAL;
	XSYNCOUTKEEPPOSITION : BOOL;
END_VAR
VAR_OUTPUT
	XSYNCOUTDONE : BOOL;
END_VAR
VAR_IN_OUT
	AXESGROUP : AXES_GROUP_KIN;
	FBBASE : L_MC4P_Template_AG_KIN;
END_VAR
END_METHOD

METHOD SYNCHRON : BOOL
VAR_INPUT
	PASCCNVVALUESCCS : POINTER TO ARRAY [1..6] OF L_MC4P_AxisProfile;
	PTRAFO_BASE_MCS : POINTER TO L_MC4P_CoordTrafo;
END_VAR
END_METHOD

METHOD STATE_AGSTOP
VAR_INPUT
	XEXECUTE : BOOL;
END_VAR
VAR_IN_OUT
	AXESGROUP : AXES_GROUP_KIN;
	FBBASE : L_MC4P_Template_AG_KIN;
END_VAR
END_METHOD

METHOD STATE_ABORTING
VAR_INPUT
	XEXECUTE : BOOL;
END_VAR
VAR_IN_OUT
	AXESGROUP : AXES_GROUP_KIN;
	FBBASE : L_MC4P_Template_AG_KIN;
END_VAR
END_METHOD

METHOD STATE_ERROR
VAR_INPUT
	XEXECUTE : BOOL;
END_VAR
VAR_IN_OUT
	AXESGROUP : AXES_GROUP_KIN;
	FBBASE : L_MC4P_Template_AG_KIN;
END_VAR
END_METHOD

METHOD STATE_INITIAL
VAR_INPUT
	XEXECUTE : BOOL;
	XSETDYNPCSINDEPENDANT : BOOL;
END_VAR
VAR_IN_OUT
	AXESGROUP : AXES_GROUP_KIN;
	FBBASE : L_MC4P_Template_AG_KIN;
END_VAR
END_METHOD

METHOD STATE_SYNCIN
VAR_INPUT
	XEXECUTE : BOOL;
END_VAR
VAR_IN_OUT
	AXESGROUP : AXES_GROUP_KIN;
	FBBASE : L_MC4P_Template_AG_KIN;
END_VAR
END_METHOD

METHOD STATE_SYNCOUT
VAR_INPUT
	XEXECUTE : BOOL;
	XABORT : BOOL;
END_VAR
VAR_IN_OUT
	AXESGROUP : AXES_GROUP_KIN;
	FBBASE : L_MC4P_Template_AG_KIN;
END_VAR
END_METHOD

METHOD STATE_SYNCHRON
VAR_INPUT
	XEXECUTE : BOOL;
END_VAR
VAR_IN_OUT
	AXESGROUP : AXES_GROUP_KIN;
	FBBASE : L_MC4P_Template_AG_KIN;
END_VAR
END_METHOD

METHOD STATE_WAITFORMOTION
VAR_INPUT
	XEXECUTE : BOOL;
END_VAR
VAR_IN_OUT
	AXESGROUP : AXES_GROUP_KIN;
	FBBASE : L_MC4P_Template_AG_KIN;
END_VAR
END_METHOD

METHOD TRACKKINEMATICS
VAR_INPUT
	XEXECUTE : BOOL;
	XABORT : BOOL;
	XSETDYNPCSINDEPENDANT : BOOL;
END_VAR
VAR_IN_OUT
	AXESGROUP : AXES_GROUP_KIN;
	FBBASE : L_MC4P_Template_AG_KIN;
END_VAR
END_METHOD

(* ---- L_MC4P_TRAFOEXTENSIONBASE.fb ---- *)
FUNCTION_BLOCK L_MC4P_TRAFOEXTENSIONBASE EXTENDS L_MC4P_Template_AG_KIN
END_FUNCTION_BLOCK

METHOD BACKWARDTRANSFORMATIONEXTENSION : L_IE1P_Error
VAR_INPUT
	PAXES_POS : POINTER TO ARRAY [1..6] OF LREAL;
	PJOINT_POS : POINTER TO ARRAY [1..6] OF LREAL;
END_VAR
END_METHOD

METHOD CHECKINPUTS : L_IE1P_Error
VAR_IN_OUT
	AXESGROUP : AXES_GROUP_KIN;
END_VAR
END_METHOD

METHOD FORWARDTRANSFORMATIONEXTENSION : L_IE1P_Error
VAR_INPUT
	PAXES_POS : POINTER TO ARRAY [1..6] OF LREAL;
	PJOINT_POS : POINTER TO ARRAY [1..6] OF LREAL;
END_VAR
END_METHOD

METHOD GENERALIZEDFORCE_ACS2JCS : L_IE1P_Error
VAR_INPUT
	PAXES_FORCE : POINTER TO ARRAY [1..6] OF LREAL;
	PJOINT_FORCE : POINTER TO ARRAY [1..6] OF LREAL;
END_VAR
END_METHOD

METHOD GENERALIZEDFORCE_JCS2ACS : L_IE1P_Error
VAR_INPUT
	PAXES_FORCE : POINTER TO ARRAY [1..6] OF LREAL;
	PJOINT_FORCE : POINTER TO ARRAY [1..6] OF LREAL;
END_VAR
END_METHOD

(* ---- L_MC4P_TRAFOINFO.fb ---- *)
FUNCTION_BLOCK L_MC4P_TRAFOINFO
VAR_INPUT
	ALITURNS : ARRAY [1..6] OF LINT;
	AIQUADRANT : ARRAY [1..6] OF INT;
	AICONFIG : ARRAY [1..6] OF INT;
	XCHECKQUADRANT : BOOL;
	ALRNEIGHBOUR : ARRAY [1..6] OF LREAL;
	ICHECKNEIGHBOURHOOD : INT;
	ETOOLSYSTEM : L_MC4P_ToolSystem;
END_VAR
VAR
	TYPEID : L_MC4P_KinematicType;
END_VAR
END_FUNCTION_BLOCK

METHOD COPYFROM : L_IE1P_Error
VAR_INPUT
	SCSOURCE : REFERENCE TO L_MC4P_TrafoInfo;
END_VAR
END_METHOD

METHOD FB_INIT : BOOL
VAR_INPUT
	BINITRETAINS : BOOL;
	BINCOPYCODE : BOOL;
END_VAR
END_METHOD

METHOD RESET
END_METHOD

(* ---- L_MC4P_VIRTUALTIME.fb ---- *)
FUNCTION_BLOCK L_MC4P_VIRTUALTIME
VAR_INPUT
	XENABLE : BOOL;
	LRCYCLETIME : LREAL;
	LROVRREQUESTED : LREAL := 1.0;
END_VAR
VAR_OUTPUT
	LRVIRTUALTIMECYCLE : LREAL;
	LROVRACTUAL : LREAL;
	LRDOVRACTUAL : LREAL;
	XERROR : BOOL := FALSE;
	EERRORID : L_IE1P_Error;
END_VAR
VAR
	_REFTIMEFILTER : REFERENCE TO L_USPP_Filter;
	_FBPT2 : L_USPP_PT2Filter;
	_XTIMEFILTERDONE : BOOL;
	_XPAUSE : BOOL := FALSE;
	_XFORCEOVREQ1 : BOOL := FALSE;
	XPAUSE : BOOL;
END_VAR
END_FUNCTION_BLOCK

METHOD CALLTIMEFILTER
END_METHOD

METHOD ENTRYCYCLE
END_METHOD

METHOD FORCESTOPOVREQ1
END_METHOD

METHOD IDENTIFYTIMEFILTER : BOOL
VAR_INPUT
	FBTIMEFILTER : REFERENCE TO L_USPP_Filter;
END_VAR
END_METHOD

METHOD LEAVECYCLE
END_METHOD

METHOD REPLACETIMEFILTER
VAR_INPUT
	FBTIMEFILTER : REFERENCE TO L_USPP_Filter;
END_VAR
END_METHOD

METHOD FB_INIT : BOOL
VAR_INPUT
	BINITRETAINS : BOOL;
	BINCOPYCODE : BOOL;
END_VAR
END_METHOD

(* ---- L_MC4P_VISU_AXES_GROUP_KIN.fb ---- *)
FUNCTION_BLOCK L_MC4P_VISU_AXES_GROUP_KIN
VAR_INPUT
	M_INPUT_INST_STR : STRING;
	XENABLEVISU : BOOL := FALSE;
	XTEST : BOOL := FALSE;
	XSHOWPATH : BOOL := TRUE;
	PAXESGROUP : POINTER TO AXES_GROUP_KIN;
END_VAR
VAR
	FBKINCOORDPROVIDER : L_MC4P_KinCoordProvider;
	XENABLEVISUOLD : BOOL := FALSE;
	ALRACSTESTPOS : ARRAY [1..6] OF LREAL := [6(0)];
	ALRACSPOS : ARRAY [1..6] OF LREAL := [6(0)];
	ALRJCSPOS : ARRAY [1..6] OF LREAL := [6(0)];
	ALRXTCS_MCS : ARRAY [1..6] OF LREAL := [6(0)];
	ALRXTCS_WCS : ARRAY [1..6] OF LREAL := [6(0)];
	ALRXEE_MCS : ARRAY [1..6] OF LREAL := [6(0)];
	ALRMCS_WCS : ARRAY [1..6] OF LREAL := [6(0)];
	ALRWCS_MCS : ARRAY [1..6] OF LREAL := [6(0)];
	COORDTMP : MC_COORD_REF;
	AXDISPLAYINVISIBLE : ARRAY [1..12] OF BOOL;
	AXDISPLAYINACTIVE : ARRAY [1..12] OF BOOL;
	XSHOWCONFIGELEMENTS : BOOL := FALSE;
	IDX : INT;
	XINIT : BOOL := TRUE;
	XREINIT : BOOL := TRUE;
	EKINEMATIC : L_MC4P_KinematicType := L_MC4P_KinematicType.NoKinematic;
	XSCALING : BOOL;
	FRAMELIMITATION : ARRAY [1..6] OF LREAL;
	XSHOWFRAME : BOOL := FALSE;
	XRECALCSCALINGS : BOOL := FALSE;
	XVISUPCSACTIVE : BOOL := FALSE;
	LRUNITSTOPIXELFRAME1 : LREAL := 1;
	LRUNITSTOPIXELFRAME2 : LREAL := 1;
	LRMCS0FRAME1 : ARRAY [1..2] OF LREAL := [200, 200];
	LRMCS0FRAME2 : ARRAY [1..2] OF LREAL := [50, 350];
	ALRRTCS2MCS : ARRAY [1..3, 1..3] OF LREAL;
	ALRRMCS2TCS : ARRAY [1..3, 1..3] OF LREAL;
	ALRRMCS2FRAME1 : ARRAY [1..3, 1..3] OF LREAL;
	ALRRFRAME12MCS : ARRAY [1..3, 1..3] OF LREAL;
	ALRRMCS2FRAME2 : ARRAY [1..3, 1..3] OF LREAL;
	ALRRFRAME22MCS : ARRAY [1..3, 1..3] OF LREAL;
	ALRRTCS2FRAME1 : ARRAY [1..3, 1..3] OF LREAL;
	ALRRTCS2FRAME2 : ARRAY [1..3, 1..3] OF LREAL;
	ALRRWCS2FRAME1 : ARRAY [1..3, 1..3] OF LREAL;
	ALRRWCS2FRAME2 : ARRAY [1..3, 1..3] OF LREAL;
	ALRRWCS2MCS : ARRAY [1..3, 1..3] OF LREAL;
	ALRRMCS2WCS : ARRAY [1..3, 1..3] OF LREAL;
	ALRXWCSFRAME1 : ARRAY [1..4] OF LREAL;
	ALRYWCSFRAME1 : ARRAY [1..4] OF LREAL;
	ALRZWCSFRAME1 : ARRAY [1..4] OF LREAL;
	ALRXWCSFRAME2 : ARRAY [1..4] OF LREAL;
	ALRYWCSFRAME2 : ARRAY [1..4] OF LREAL;
	ALRZWCSFRAME2 : ARRAY [1..4] OF LREAL;
	ALRXMCSFRAME1 : ARRAY [1..4] OF LREAL;
	ALRYMCSFRAME1 : ARRAY [1..4] OF LREAL;
	ALRZMCSFRAME1 : ARRAY [1..4] OF LREAL;
	ALRXMCSFRAME2 : ARRAY [1..4] OF LREAL;
	ALRYMCSFRAME2 : ARRAY [1..4] OF LREAL;
	ALRZMCSFRAME2 : ARRAY [1..4] OF LREAL;
	ALRXTCSFRAME1 : ARRAY [1..4] OF LREAL;
	ALRYTCSFRAME1 : ARRAY [1..4] OF LREAL;
	ALRZTCSFRAME1 : ARRAY [1..4] OF LREAL;
	ALRXTCSFRAME2 : ARRAY [1..4] OF LREAL;
	ALRYTCSFRAME2 : ARRAY [1..4] OF LREAL;
	ALRZTCSFRAME2 : ARRAY [1..4] OF LREAL;
	ALRPATH_MCS : ARRAY [1..100, 1..3] OF LREAL;
	ALRPATH_FRAME1 : ARRAY [1..100, 1..2] OF LREAL;
	ALRPATH_FRAME2 : ARRAY [1..100, 1..2] OF LREAL;
	XRESETPATHARRAY : BOOL := TRUE;
	ALRXTMP : ARRAY [1..3] OF LREAL;
	LRANGLEX : LREAL;
	LRANGLEY : LREAL;
	LRANGLEZ : LREAL;
	LRPROJLENGTHX : LREAL;
	LRPROJLENGTHY : LREAL;
	LRPROJLENGTHZ : LREAL;
	LRROTZ_FRAME1DEG : LREAL := 0;
	LRROTZ_FRAME1OLDDEG : LREAL := 0;
	LRROTZ_FRAME2DEG : LREAL := 0;
	LRROTZ_FRAME2OLDDEG : LREAL := 0;
	LRVALIDCOLOR : LREAL;
	ETRAFOERROR : L_IE1P_Error;
	XVALID : BOOL := FALSE;
	WSELECTFRAME1 : WORD;
	WSELECTFRAME2 : WORD;
	WSELECTFRAME1OLD : WORD;
	WSELECTFRAME2OLD : WORD;
	IFELD : INT := 1;
	USICOUNTERVAL : USINT := 0;
	AXSHOWPCS : ARRAY [1..16] OF BOOL;
	ALRPCSPOS_WCS : ARRAY [1..16, 1..6] OF LREAL;
	ALRRPCS2MCS : ARRAY [1..3, 1..3] OF LREAL;
	ALRRMCS2PCS : ARRAY [1..3, 1..3] OF LREAL;
	ALRRPCS2FRAME1 : ARRAY [1..3, 1..3] OF LREAL;
	ALRRPCS2FRAME2 : ARRAY [1..3, 1..3] OF LREAL;
	ALRXPCSFRAME1 : ARRAY [1..4] OF LREAL;
	ALRYPCSFRAME1 : ARRAY [1..4] OF LREAL;
	ALRZPCSFRAME1 : ARRAY [1..4] OF LREAL;
	ALRXPCSFRAME2 : ARRAY [1..4] OF LREAL;
	ALRYPCSFRAME2 : ARRAY [1..4] OF LREAL;
	ALRZPCSFRAME2 : ARRAY [1..4] OF LREAL;
	ALRMCS_T_WCS : ARRAY [1..4, 1..4] OF LREAL;
	ALRMCS_T_PCS : ARRAY [1..4, 1..4] OF LREAL;
	ALRWCS_T_PCS : ARRAY [1..4, 1..4] OF LREAL;
	XSHOWPCS : BOOL := FALSE;
	ESHOWPCS : L_MC4P_CoordSystem := L_MC4P_CoordSystem.PCS_1;
	XVISUHASPARAMETER : BOOL := FALSE;
	XSHOWMCS : BOOL := TRUE;
	XSHOWWCS : BOOL := FALSE;
	USIPATHCYCLES : USINT := 10;
	HEVENTCOMMCYCLE : Systypes.RTS_IEC_HANDLE := SysTypes.RTS_INVALID_HANDLE;
	HINTERFACECOMMCYCLE : Systypes.RTS_IEC_HANDLE := SysTypes.RTS_INVALID_HANDLE;
	ITFCALLBACK : CmpEventMgr.ICmpEventCallback;
	DWEVENTCOUNTER : DWORD;
	LRMCSPIXEL : LREAL := 50;
	LRTCSPIXEL : LREAL := 30;
	LRWCSPIXEL : LREAL := 50;
END_VAR
END_FUNCTION_BLOCK

METHOD COMMONINITIALIZE
END_METHOD

METHOD COMMONMAIN
END_METHOD

METHOD COORDSYSFRAME1
END_METHOD

METHOD COORDSYSFRAME2
END_METHOD

METHOD FB_EXIT : BOOL
VAR_INPUT
	BINCOPYCODE : BOOL;
END_VAR
END_METHOD

METHOD INITIALIZE
END_METHOD

METHOD KINEMATICFRAME1
END_METHOD

METHOD KINEMATICFRAME2
END_METHOD

METHOD PATH
END_METHOD

METHOD PATHFRAME1
END_METHOD

METHOD PATHFRAME2
END_METHOD

METHOD RECALCSCALINGS
END_METHOD

METHOD UPDATEORIENTATIONFRAME1
END_METHOD

METHOD UPDATEORIENTATIONFRAME2
END_METHOD

METHOD FB_INIT : BOOL
VAR_INPUT
	BINITRETAINS : BOOL;
	BINCOPYCODE : BOOL;
END_VAR
END_METHOD

METHOD EVENTCALLBACK : UDINT
VAR_INPUT
	PEVENTPARAM : POINTER TO EventParam;
END_VAR
END_METHOD

METHOD REGISTEREVENT
END_METHOD

METHOD UNREGISTEREVENT
END_METHOD

(* ---- L_MC4P_WRITEBOOLPARAMETER.fb ---- *)
FUNCTION_BLOCK L_MC4P_WRITEBOOLPARAMETER EXTENDS L_MC4P_Template_AG_KIN
VAR_INPUT
	XEXECUTE : BOOL;
	DIPARAMETERNUMBER : DINT;
	XVALUE : BOOL;
END_VAR
VAR_OUTPUT
	XDONE : BOOL;
	XBUSY : BOOL;
	XERROR : BOOL;
	EERRORID : L_IE1P_Error;
END_VAR
VAR
	XEXECUTEOLD : BOOL := FALSE;
	XRESETOUTPUT : BOOL := FALSE;
	WERRORID_INT : WORD;
END_VAR
END_FUNCTION_BLOCK

METHOD FB_RESET : BOOL
END_METHOD

(* ---- L_MC4P_WRITEPARAMETER.fb ---- *)
FUNCTION_BLOCK L_MC4P_WRITEPARAMETER EXTENDS L_MC4P_Template_AG_KIN
VAR_INPUT
	XEXECUTE : BOOL;
	DIPARAMETERNUMBER : DINT;
	LRVALUE : LREAL;
END_VAR
VAR_OUTPUT
	XDONE : BOOL;
	XBUSY : BOOL;
	XERROR : BOOL;
	EERRORID : L_IE1P_Error;
END_VAR
VAR
	XEXECUTEOLD : BOOL := FALSE;
	XRESETOUTPUT : BOOL := FALSE;
	WERRORID_INT : WORD;
END_VAR
END_FUNCTION_BLOCK

METHOD FB_RESET : BOOL
END_METHOD

(* ---- L_MC4P_WRITEPATHFILE_INTERNAL.fb ---- *)
FUNCTION_BLOCK L_MC4P_WRITEPATHFILE_INTERNAL
VAR_INPUT
	XEXECUTE : BOOL;
	SFILENAME : STRING;
	SFILEADRES : STRING := '\USBStorage\IPC\PLC\MovePathData\';
	DINUMOFLINES : DINT := 200;
END_VAR
VAR_OUTPUT
	XDONE : BOOL;
	XBUSY : BOOL;
	XCOMMANDABORTED : BOOL;
	XERROR : BOOL;
	EERRORID : L_IE1P_Error;
END_VAR
VAR_IN_OUT
	ASPATHFILE : ARRAY [1..200] OF STRING(255);
END_VAR
VAR
	WSTATE : WORD;
	XNEWFILE_INT : BOOL;
	DILINENO_INT : DINT;
	DINUMOFLINES_INT : DINT;
	UDIPOSINFILE : UDINT;
	FB_SEMA : L_MC1P_CriticalSection;
	REQUESTSINFO : DWORD;
	REQUESTSINFO_OLD : DWORD;
	DWRTRIG : DWORD;
	DWFTRIG : DWORD;
	SFILE_INT : STRING := '';
	WTASKCYCLECOUNTER : WORD := 0;
	XLOWTASKBUSY_INT : BOOL;
	XLOWTASKDONE_INT : BOOL;
	XLOWTASKERROR_INT : BOOL;
	ELOWTASKERRORID_INT : L_IE1P_Error;
	RES : SYSFILE.RTS_IEC_ResULT;
	HFILE : SYSFILE.RTS_IEC_HANDLE;
	UDILENGTHFILE : UDINT;
	UDIFSIZE : UDINT;
	XTESTINMOTIONTASK : BOOL := FALSE;
	ILINELEN_INT : INT;
	XERROR_TIMEOUT : BOOL;
	FILDCR : FILE.DirCreate;
	SLINE : STRING(255);
	XDECODEINMOTIONTASK : BOOL;
END_VAR
END_FUNCTION_BLOCK

METHOD ABORTFB : UDINT
END_METHOD

METHOD CALL_ERRORHANDLER
END_METHOD

METHOD CALL_FBMETHODS
END_METHOD

METHOD CALL_OUTPUT
END_METHOD

METHOD CALL_REQUESTS_EXT
END_METHOD

METHOD CALL_RESETCOMMANDS
END_METHOD

METHOD CALL_RESETOUTPUT
END_METHOD

METHOD CALL_STATEMACHINE
END_METHOD

METHOD RESETREADDATA
END_METHOD

METHOD CALL_WRITEFILE
END_METHOD

METHOD EXECUTEFREERUNTASK
END_METHOD

METHOD MAIN
END_METHOD

METHOD ABORT : UDINT
END_METHOD

METHOD EXECUTE : UDINT
END_METHOD

(* ---- MC_ADDAXISTOGROUP.fb ---- *)
FUNCTION_BLOCK MC_ADDAXISTOGROUP EXTENDS L_MC4P_Template_AG_KIN
VAR_INPUT
	EXECUTE : BOOL;
	IDENTINGROUP : IDENT_IN_GROUP_REF;
END_VAR
VAR_OUTPUT
	DONE : BOOL;
	BUSY : BOOL;
	ERROR : BOOL;
	ERRORID : L_IE1P_Error;
END_VAR
VAR_IN_OUT
	AXIS : AXIS_REF;
END_VAR
VAR
	XERRORINTERN : BOOL;
	EERRORIDINTERN : L_IE1P_Error := L_IE1P_Error.NoError;
	XEXECUTEOLD : BOOL;
	XRESETOUTPUT : BOOL;
	PSDUMMY : POINTER TO STRING;
	PAXIS : POINTER TO POINTER TO AXIS_REF;
END_VAR
END_FUNCTION_BLOCK

(* ---- MC_GROUPDISABLE.fb ---- *)
FUNCTION_BLOCK MC_GROUPDISABLE EXTENDS L_MC4P_Template_AG_REF
VAR_INPUT
	EXECUTE : BOOL;
END_VAR
VAR_OUTPUT
	DONE : BOOL;
	BUSY : BOOL;
	ERROR : BOOL;
	ERRORID : L_IE1P_Error;
END_VAR
VAR
	XEXECUTEOLD : BOOL;
	IDX : WORD;
	XRESETOUTPUT : BOOL;
	XVIRTAXISENABLED : BOOL;
	PXDUMMY : POINTER TO BOOL;
	PAXESGROUP : POINTER TO AXES_GROUP_KIN;
	WDISABLECNTR : WORD;
	WDISABLECNTRMAX : WORD := 50;
	XREADYFORDISABLE : BOOL;
	WSTATE : WORD;
	XDOWHILE : BOOL;
	ICNT : INT;
END_VAR
END_FUNCTION_BLOCK

(* ---- MC_GROUPENABLE.fb ---- *)
FUNCTION_BLOCK MC_GROUPENABLE EXTENDS L_MC4P_Template_AG_REF
VAR_INPUT
	EXECUTE : BOOL;
END_VAR
VAR_OUTPUT
	DONE : BOOL;
	BUSY : BOOL;
	ERROR : BOOL;
	ERRORID : L_IE1P_Error;
END_VAR
VAR
	XEXECUTEOLD : BOOL;
	IDX : WORD;
	XRESETOUTPUT : BOOL;
	XREALAXISENABLED : BOOL;
	XREALAXISSTANDSTILL : BOOL;
	XVIRTAXISENABLED : BOOL;
	WSTEP : WORD;
	PXDUMMY : POINTER TO BOOL;
	ALRKARTPOS : ARRAY [1..6] OF LREAL;
	ALRACTAXESPOS : ARRAY [1..6] OF LREAL;
	ALRCALCULATEDAXESPOS : ARRAY [1..6] OF LREAL;
	ALRAXESPOSDIFF : ARRAY [1..6] OF LREAL;
	PAXESGROUP : POINTER TO AXES_GROUP_KIN;
	XERRORINTERN : BOOL;
	EERRORIDINTERN : L_IE1P_Error;
	EERRORIDINTERN2 : L_IE1P_Error;
	SCERROR : L_MC4P_ErrorStruct;
	SCINFO : L_MC4P_TrafoInfo;
END_VAR
END_FUNCTION_BLOCK

METHOD FB_INIT : BOOL
VAR_INPUT
	BINITRETAINS : BOOL;
	BINCOPYCODE : BOOL;
END_VAR
END_METHOD

(* ---- MC_GROUPHOME.fb ---- *)
FUNCTION_BLOCK MC_GROUPHOME EXTENDS L_MC4P_Template_AG_KIN_Licence
VAR_INPUT
	EXECUTE : BOOL;
	POSITION : ARRAY [1..12] OF LREAL;
	HOMINGORDER : ARRAY [1..12] OF L_MC4P_HomingOrder := [12(0)];
	HOMEABSSWITCH : ARRAY [1..12] OF BOOL;
	USEEXTPARAMETER : ARRAY [1..12] OF BOOL;
	EXTPARAMETER : ARRAY [1..12] OF L_MC1P_HomeParameter;
	EXTTP : ARRAY [1..12] OF MC_TRIGGER_REF;
END_VAR
VAR_OUTPUT
	DONE : BOOL;
	BUSY : BOOL;
	ACTIVE : BOOL;
	COMMANDABORTED : BOOL;
	ERROR : BOOL;
	ERRORID : L_IE1P_Error;
	AXISDONE : ARRAY [1..12] OF BOOL;
END_VAR
VAR
	HOME : L_MC4P_GroupHome_Internal;
END_VAR
END_FUNCTION_BLOCK

(* ---- MC_GROUPREADACTUALACCELERATION.fb ---- *)
FUNCTION_BLOCK MC_GROUPREADACTUALACCELERATION EXTENDS L_MC4P_Template_AG_KIN
VAR_INPUT
	ENABLE : BOOL;
	COORDSYSTEM : L_MC4P_CoordSystem;
END_VAR
VAR_OUTPUT
	VALID : BOOL;
	BUSY : BOOL;
	ERROR : BOOL;
	ERRORID : L_IE1P_Error;
	ACCELERATION : ARRAY [1..12] OF LREAL;
	PATHACCELERATION : LREAL;
END_VAR
VAR
	IDX : WORD;
	XENABLEOLD : BOOL;
	PCOORDTRAFO : POINTER TO L_MC4P_CoordTrafo;
	ALRACCELERATIONTMP1 : ARRAY [1..6] OF LREAL;
	ALRACCELERATIONTMP2 : ARRAY [1..6] OF LREAL;
	ALRVELOCITYTMP1 : ARRAY [1..6] OF LREAL;
	ALRVELOCITYTMP2 : ARRAY [1..6] OF LREAL;
	ALRPOSITIONTMP : ARRAY [1..6] OF LREAL;
	ALRPOSVEKPCS2TCS : ARRAY [1..3] OF LREAL;
	ROT_MAT : ARRAY [1..3, 1..3] OF LREAL;
	ROT_MATT : ARRAY [1..3, 1..3] OF LREAL;
	ALRTMP : ARRAY [1..3] OF LREAL;
	T1 : LREAL;
	T5 : LREAL;
	T6 : LREAL;
	T7 : LREAL;
	T13 : LREAL;
	T20 : LREAL;
	T21 : LREAL;
	T26 : LREAL;
	X : LREAL;
	Y : LREAL;
	XPUNKT : LREAL;
	YPUNKT : LREAL;
	XPUNKTPUNKT : LREAL;
	YPUNKTPUNKT : LREAL;
END_VAR
END_FUNCTION_BLOCK

(* ---- MC_GROUPREADACTUALPOSITION.fb ---- *)
FUNCTION_BLOCK MC_GROUPREADACTUALPOSITION EXTENDS L_MC4P_Template_AG_KIN
VAR_INPUT
	ENABLE : BOOL;
	COORDSYSTEM : L_MC4P_CoordSystem;
END_VAR
VAR_OUTPUT
	VALID : BOOL;
	BUSY : BOOL;
	ERROR : BOOL;
	ERRORID : L_IE1P_Error;
	POSITION : ARRAY [1..12] OF LREAL;
END_VAR
VAR
	XUSESETVALUES : BOOL := FALSE;
	READPOSITION : L_MC4P_GroupReadActualPosition_Internal;
	USESETVALUES : BOOL;
END_VAR
END_FUNCTION_BLOCK

(* ---- MC_GROUPREADACTUALVELOCITY.fb ---- *)
FUNCTION_BLOCK MC_GROUPREADACTUALVELOCITY EXTENDS L_MC4P_Template_AG_KIN
VAR_INPUT
	ENABLE : BOOL;
	COORDSYSTEM : L_MC4P_CoordSystem;
END_VAR
VAR_OUTPUT
	VALID : BOOL;
	BUSY : BOOL;
	ERROR : BOOL;
	ERRORID : L_IE1P_Error;
	VELOCITY : ARRAY [1..12] OF LREAL;
	PATHVELOCITY : LREAL;
END_VAR
VAR
	XUSESETVALUES : BOOL := FALSE;
	READVEL : L_MC4P_GroupReadActualVelocity_Internal;
	USESETVALUES : BOOL;
END_VAR
END_FUNCTION_BLOCK

(* ---- MC_GROUPREADERROR.fb ---- *)
FUNCTION_BLOCK MC_GROUPREADERROR EXTENDS L_MC4P_Template_AG_REF
VAR_INPUT
	ENABLE : BOOL;
END_VAR
VAR_OUTPUT
	VALID : BOOL;
	BUSY : BOOL;
	ERROR : BOOL;
	ERRORID : L_IE1P_Error;
	GROUPWARNING : BOOL;
	GROUPERROR : BOOL;
	GROUPERRORID : L_IE1P_Error;
	PINSTANCENAME : POINTER TO STRING := ADR(NoError);
	TIMESTAMP : TIME;
END_VAR
VAR
	XENABLEOLD : BOOL;
	NOERROR : STRING := '';
END_VAR
END_FUNCTION_BLOCK

(* ---- MC_GROUPREADSTATUS.fb ---- *)
FUNCTION_BLOCK MC_GROUPREADSTATUS EXTENDS L_MC4P_Template_AG_KIN
VAR_INPUT
	ENABLE : BOOL;
END_VAR
VAR_OUTPUT
	VALID : BOOL;
	BUSY : BOOL;
	ERROR : BOOL;
	ERRORID : L_IE1P_Error;
	GROUPMOVING : BOOL;
	GROUPHOMING : BOOL;
	GROUPERRORSTOP : BOOL;
	GROUPSTANDBY : BOOL;
	GROUPSTOPPING : BOOL;
	GROUPDISABLED : BOOL;
	CONSTANTVELOCITY : BOOL;
	ACCELERATING : BOOL;
	DECELERATING : BOOL;
	INPOSITION : BOOL;
	STANDSTILL : BOOL;
END_VAR
VAR
	READSTATUS : L_MC4P_GroupReadStatus_Internal;
END_VAR
END_FUNCTION_BLOCK

(* ---- MC_GROUPRESET.fb ---- *)
FUNCTION_BLOCK MC_GROUPRESET EXTENDS L_MC4P_Template_AG_REF
VAR_INPUT
	EXECUTE : BOOL;
END_VAR
VAR_OUTPUT
	DONE : BOOL;
	BUSY : BOOL;
	ERROR : BOOL;
	ERRORID : L_IE1P_Error;
END_VAR
VAR
	GROUPRESET : L_MC4P_GroupReset_Internal;
END_VAR
END_FUNCTION_BLOCK

(* ---- MC_GROUPSETPOSITION.fb ---- *)
FUNCTION_BLOCK MC_GROUPSETPOSITION EXTENDS L_MC4P_Template_AG_KIN
VAR_INPUT
	EXECUTE : BOOL;
	POSITION : ARRAY [1..12] OF LREAL;
	RELATIVE : BOOL := FALSE;
END_VAR
VAR_OUTPUT
	DONE : BOOL;
	BUSY : BOOL;
	ACTIVE : BOOL;
	ERROR : BOOL;
	ERRORID : L_IE1P_Error;
END_VAR
VAR
	SETPOSITION : L_MC4P_GroupSetPosition_Internal;
END_VAR
END_FUNCTION_BLOCK

(* ---- MC_GROUPSTOP.fb ---- *)
FUNCTION_BLOCK MC_GROUPSTOP EXTENDS L_MC4P_Template_AG_KIN_Licence
VAR_INPUT
	EXECUTE : BOOL;
	DECELERATION : LREAL;
	JERK : LREAL;
END_VAR
VAR_OUTPUT
	DONE : BOOL;
	BUSY : BOOL;
	ACTIVE : BOOL;
	COMMANDABORTED : BOOL;
	ERROR : BOOL;
	ERRORID : L_IE1P_Error;
END_VAR
VAR
	STOP : L_MC4P_GroupStop_Internal;
END_VAR
END_FUNCTION_BLOCK

(* ---- MC_MOVECIRCULARABSOLUTE.fb ---- *)
FUNCTION_BLOCK MC_MOVECIRCULARABSOLUTE EXTENDS L_MC4P_Template_MoveLicence
VAR_INPUT
	EXECUTE : BOOL;
	CIRCMODE : L_MC4P_CircMode;
	AUXPOINT : ARRAY [1..12] OF LREAL;
	ENDPOINT : ARRAY [1..12] OF LREAL;
	PATHCHOICE : MC_CIRC_PATHCHOICE;
	VELOCITY : LREAL;
	ACCELERATION : LREAL;
	DECELERATION : LREAL;
	JERK : LREAL;
	COORDSYSTEM : L_MC4P_CoordSystem;
	BUFFERMODE : MC_BUFFER_MODE;
	TRANSITIONMODE : MC_TRANSITION_MODE;
	TRANSITIONPARAMETER : ARRAY [1..12] OF LREAL := [12(0)];
	AEAUXMODE : ARRAY [1..6] OF L_MC4P_AuxMode;
	ORIENTATIONMODE : L_MC4P_Orientation_Mode := L_MC4P_Orientation_Mode.ShortestSpacialWay;
	DIRECTION : ARRAY [4..6] OF MC_DIRECTION := [3(MC_DIRECTION.mcShortestWay)];
END_VAR
VAR_OUTPUT
	DONE : BOOL;
	BUSY : BOOL;
	ACTIVE : BOOL;
	COMMANDABORTED : BOOL;
	ERROR : BOOL;
	ERRORID : L_IE1P_Error;
END_VAR
VAR
	MOVECIRC : L_MC4P_MoveCircularAbsolute_Internal;
	PMOVE : POINTER TO L_MC4P_MoveContPath;
END_VAR
END_FUNCTION_BLOCK

(* ---- MC_MOVECIRCULARRELATIVE.fb ---- *)
FUNCTION_BLOCK MC_MOVECIRCULARRELATIVE EXTENDS L_MC4P_Template_MoveLicence
VAR_INPUT
	EXECUTE : BOOL;
	CIRCMODE : L_MC4P_CircMode;
	AUXPOINT : ARRAY [1..12] OF LREAL;
	ENDPOINT : ARRAY [1..12] OF LREAL;
	PATHCHOICE : MC_CIRC_PATHCHOICE;
	VELOCITY : LREAL;
	ACCELERATION : LREAL;
	DECELERATION : LREAL;
	JERK : LREAL;
	COORDSYSTEM : L_MC4P_CoordSystem;
	BUFFERMODE : MC_BUFFER_MODE;
	TRANSITIONMODE : MC_TRANSITION_MODE;
	TRANSITIONPARAMETER : ARRAY [1..12] OF LREAL := [12(0)];
	AEAUXMODE : ARRAY [1..6] OF L_MC4P_AuxMode;
	ORIENTATIONMODE : L_MC4P_Orientation_Mode := L_MC4P_Orientation_Mode.ShortestSpacialWay;
	DIRECTION : ARRAY [4..6] OF MC_DIRECTION := [3(MC_DIRECTION.mcShortestWay)];
END_VAR
VAR_OUTPUT
	DONE : BOOL;
	BUSY : BOOL;
	ACTIVE : BOOL;
	COMMANDABORTED : BOOL;
	ERROR : BOOL;
	ERRORID : L_IE1P_Error;
END_VAR
VAR
	MOVECIRC : L_MC4P_MoveCircularRelative_Internal;
	PMOVE : POINTER TO L_MC4P_MoveContPath;
END_VAR
END_FUNCTION_BLOCK

(* ---- MC_MOVEDIRECTABSOLUTE.fb ---- *)
FUNCTION_BLOCK MC_MOVEDIRECTABSOLUTE EXTENDS L_MC4P_Template_MoveLicence
VAR_INPUT
	EXECUTE : BOOL;
	POSITION : ARRAY [1..12] OF LREAL;
	COORDSYSTEM : L_MC4P_CoordSystem;
	BUFFERMODE : MC_BUFFER_MODE;
	TRANSITIONMODE : MC_TRANSITION_MODE;
	TRANSITIONPARAMETER : ARRAY [1..12] OF LREAL := [12(0)];
	AITARGETCONFIGURATION : ARRAY [1..6] OF INT;
	DIRECTION : ARRAY [1..6] OF MC_DIRECTION := [6(MC_DIRECTION.mcShortestWay)];
END_VAR
VAR_OUTPUT
	DONE : BOOL;
	BUSY : BOOL;
	ACTIVE : BOOL;
	COMMANDABORTED : BOOL;
	ERROR : BOOL;
	ERRORID : L_IE1P_Error;
END_VAR
VAR
	MOVEDIRECT : L_MC4P_MoveDirectAbsolute_Internal;
	PMOVE : POINTER TO L_MC4P_MoveContPath;
END_VAR
END_FUNCTION_BLOCK

(* ---- MC_MOVEDIRECTRELATIVE.fb ---- *)
FUNCTION_BLOCK MC_MOVEDIRECTRELATIVE EXTENDS L_MC4P_Template_MoveLicence
VAR_INPUT
	EXECUTE : BOOL;
	DISTANCE : ARRAY [1..12] OF LREAL;
	COORDSYSTEM : L_MC4P_CoordSystem;
	BUFFERMODE : MC_BUFFER_MODE;
	TRANSITIONMODE : MC_TRANSITION_MODE;
	TRANSITIONPARAMETER : ARRAY [1..12] OF LREAL := [12(0)];
	AITARGETCONFIGURATION : ARRAY [1..6] OF INT;
	DIRECTION : ARRAY [1..6] OF MC_DIRECTION := [6(MC_DIRECTION.mcShortestWay)];
END_VAR
VAR_OUTPUT
	DONE : BOOL;
	BUSY : BOOL;
	ACTIVE : BOOL;
	COMMANDABORTED : BOOL;
	ERROR : BOOL;
	ERRORID : L_IE1P_Error;
END_VAR
VAR
	MOVEDIRECT : L_MC4P_MoveDirectRelative_Internal;
	PMOVE : POINTER TO L_MC4P_MoveContPath;
END_VAR
END_FUNCTION_BLOCK

(* ---- MC_MOVELINEARABSOLUTE.fb ---- *)
FUNCTION_BLOCK MC_MOVELINEARABSOLUTE EXTENDS L_MC4P_Template_MoveLicence
VAR_INPUT
	EXECUTE : BOOL;
	POSITION : ARRAY [1..12] OF LREAL;
	VELOCITY : LREAL;
	ACCELERATION : LREAL;
	DECELERATION : LREAL;
	JERK : LREAL;
	COORDSYSTEM : L_MC4P_CoordSystem;
	BUFFERMODE : MC_BUFFER_MODE;
	TRANSITIONMODE : MC_TRANSITION_MODE;
	TRANSITIONPARAMETER : ARRAY [1..12] OF LREAL := [12(0)];
	AEAUXMODE : ARRAY [1..6] OF L_MC4P_AuxMode;
	ORIENTATIONMODE : L_MC4P_Orientation_Mode := L_MC4P_Orientation_Mode.ShortestSpacialWay;
	DIRECTION : ARRAY [4..6] OF MC_DIRECTION := [3(MC_DIRECTION.mcShortestWay)];
END_VAR
VAR_OUTPUT
	DONE : BOOL;
	BUSY : BOOL;
	ACTIVE : BOOL;
	COMMANDABORTED : BOOL;
	ERROR : BOOL;
	ERRORID : L_IE1P_Error;
END_VAR
VAR
	MOVELIN : L_MC4P_MoveLinearAbsolute_Internal;
	PMOVE : POINTER TO L_MC4P_MoveContPath;
END_VAR
END_FUNCTION_BLOCK

(* ---- MC_MOVELINEARRELATIVE.fb ---- *)
FUNCTION_BLOCK MC_MOVELINEARRELATIVE EXTENDS L_MC4P_Template_MoveLicence
VAR_INPUT
	EXECUTE : BOOL;
	DISTANCE : ARRAY [1..12] OF LREAL;
	VELOCITY : LREAL;
	ACCELERATION : LREAL;
	DECELERATION : LREAL;
	JERK : LREAL;
	COORDSYSTEM : L_MC4P_CoordSystem;
	BUFFERMODE : MC_BUFFER_MODE;
	TRANSITIONMODE : MC_TRANSITION_MODE;
	TRANSITIONPARAMETER : ARRAY [1..12] OF LREAL := [12(0)];
	AEAUXMODE : ARRAY [1..6] OF L_MC4P_AuxMode;
	ORIENTATIONMODE : L_MC4P_Orientation_Mode := L_MC4P_Orientation_Mode.ShortestSpacialWay;
	DIRECTION : ARRAY [4..6] OF MC_DIRECTION := [3(MC_DIRECTION.mcShortestWay)];
END_VAR
VAR_OUTPUT
	DONE : BOOL;
	BUSY : BOOL;
	ACTIVE : BOOL;
	COMMANDABORTED : BOOL;
	ERROR : BOOL;
	ERRORID : L_IE1P_Error;
END_VAR
VAR
	MOVELIN : L_MC4P_MoveLinearRelative_Internal;
	PMOVE : POINTER TO L_MC4P_MoveContPath;
END_VAR
END_FUNCTION_BLOCK

(* ---- MC_MOVEPATH.fb ---- *)
FUNCTION_BLOCK MC_MOVEPATH EXTENDS L_MC4P_Template_AG_KIN_Licence
VAR_INPUT
	PATHREF : MC_PATH_REF;
	EXECUTE : BOOL;
	VELOCITY : LREAL;
	ACCELERATION : LREAL;
	DECELERATION : LREAL;
	JERK : LREAL;
	COORDSYSTEM : L_MC4P_CoordSystem;
	BUFFERMODE : MC_BUFFER_MODE;
	TRANSITIONMODE : MC_TRANSITION_MODE;
	TRANSITIONPARAMETER : ARRAY [1..12] OF LREAL := [12(0)];
	MODE : WORD;
	ACKPATHHALT : BOOL;
	MACKNOWLEDGE : BOOL;
	ACKBLOCKSEARCH : BOOL;
END_VAR
VAR_OUTPUT
	DONE : BOOL;
	BUSY : BOOL;
	ACTIVE : BOOL;
	COMMANDABORTED : BOOL;
	ERROR : BOOL;
	ERRORID : L_IE1P_Error;
	SOURCELINENO : LINT;
	SOURCELINE : STRING;
	MFUNCTION : WORD;
	WAITINGFORMACKNOWLEDGE : BOOL;
	NEWVALUEMFUNCTION : BOOL;
	WAITINGFORACKPATHHALT : BOOL;
	WAITINGFORACKBLOCKSEARCH : BOOL;
END_VAR
VAR
	LRVELOCITY_INT : LREAL;
	LRACCELERATION_INT : LREAL;
	LRDECELERATION_INT : LREAL;
	LRJERK_INT : LREAL;
	ECOORDSYSTEM_INT : L_MC4P_CoordSystem;
	EBUFFERMODE_INT : MC_BUFFER_MODE;
	ETRANSITIONMODE_INT : MC_TRANSITION_MODE;
	ALRTRANSITIONPARAMETER_INT : ARRAY [1..12] OF LREAL := [12(0)];
	EMODE_INT : WORD;
	DIACKPATHHALT_INT : DINT;
	XERROR_OLD : BOOL;
	XPATHREFVALID : BOOL;
	XWPATHREFID : __XWORD;
	DWPATHREFSTATUS : DWORD;
	XPATHREFERROR : BOOL;
	XPATHREFDONE : BOOL;
	XPATHREFBUSY : BOOL;
	XPATHREFCOMMANDABORTED : BOOL;
	XPATHREFDECODING : BOOL;
	XPATHREFINTERPRETERHALT : BOOL;
	XINTERPRETERHALTACKED : BOOL;
	XPATHREFINTERPRETERHALTAPPL : BOOL;
	XPATHREFDATAACTIVE : BOOL;
	APELEMENT : ARRAY [1..GVL_MovePath.gciNumOfDecodeAsciiData] OF POINTER TO L_MC4P_Parameter_MCMove;
	PELEMENT : POINTER TO L_MC4P_Parameter_MCMove;
	SCINITELEMENT : L_MC4P_Parameter_MCMove;
	IPATHSTARTNO : INT;
	IPATHDATASIZE : UDINT;
	LIFILELINENO : LINT;
	XUPDATESOURCE : BOOL;
	XBUSY_INT : BOOL;
	XDONE_INT : BOOL;
	XCOMMANDABORTED_INT : BOOL;
	XWAITFORDONE : BOOL;
	XERROR_INT : BOOL;
	REQUESTSINFO : DWORD;
	REQUESTSINFO_OLD : DWORD;
	DWRTRIG : DWORD;
	DWFTRIG : DWORD;
	XRESETOUTPUTS : BOOL;
	XSEGMENTACTIVE_OLD : BOOL;
	MFUNCTION_OLD : WORD;
	XMACKNOWLEDGEACTIVE : BOOL;
	XSETFIRSTSOURCELINE_LOCK : BOOL;
	XWPATHREFID_LOCK : __XWORD;
	XSETPATHDATAACTIVE_LOCK : BOOL;
	XUNLOCKPATHREF : BOOL;
	DWSTATE_INT : DWORD;
	IEXECUTEELEMENTSIZE : INT;
	IEXECUTEELEMENTSIZE_LOCK : INT;
	XERRORINVALIDPATHREF : BOOL;
	XERRORPATHREFINUSE : BOOL;
	XMOVECONTPATHDONE : BOOL;
	XMOVECONTPATHBUSY : BOOL;
	XMOVECONTPATHWAITFORINTERPRETER : BOOL;
	XMOVECONTPATHCOMMANDABORTED : BOOL;
	XMOVECONTPATHCOMMANDABORTEDATHALT : BOOL;
	XMOVECONTPATHERROR : BOOL;
	EMOVECONTPATHERRORID : L_IE1P_Error;
	IACKNMOVECONTPATHNO : INT;
	FB_MOVECONTPATHCONTROL : L_MC1P_StackControlArray := STRUCT(iMaxLegth := L_MC4P_Constants.ciNumOfMoveContPath);
	XMOVECONTPATHACTIVELOCK : BOOL;
	XDISABLEMOVECONTPATH : BOOL;
	REFFBSTORE : REFERENCE TO L_MC4P_MovePathStore;
	XOPTIMISEDPATHPREPARATION_INT : BOOL := TRUE;
	IELEMENTSIZECHECKFORPROFILECALC : INT;
	INUMOFGROUPSFORCALCPROFILE : INT;
	INUMOFSEGMENTINGROUPFORCALCPROFILE : INT;
	LRTIMEGROUPFORCALCPROFILE_OLD : LREAL;
	LRTIMEGROUPFORCALCPROFILE : LREAL;
	IMAXNUMOFSEGMENTINGROUPFORCALCPROFILE : INT := 7;
	LRMAXTIMEGROUPFORCALCPROFILE : LREAL := 0.7;
	XMOTIONREQUESTED : BOOL;
	XBLOCKSEARCHACKACTIVE : BOOL;
	XBLOCKFOUND : BOOL;
	_XSEMALOCKED : BOOL;
	FBREADPOS : MC_GroupReadActualPosition;
	XOPTIMISEDPATHPREPARATION : BOOL;
END_VAR
END_FUNCTION_BLOCK

METHOD CALL_ALLOCPOINTADR
END_METHOD

METHOD CALL_DISABLEMOVECONTPATH
VAR_IN_OUT
	AXESGROUP : AXES_GROUP_KIN;
END_VAR
END_METHOD

METHOD CALL_ERRORHANDLER
VAR_IN_OUT
	AXESGROUP : AXES_GROUP_KIN;
END_VAR
END_METHOD

METHOD CALL_FBMETHODS
VAR_IN_OUT
	AXESGROUP : AXES_GROUP_KIN;
END_VAR
END_METHOD

METHOD CALL_FB_MOVECONTPATH
VAR_IN_OUT
	AXESGROUP : AXES_GROUP_KIN;
END_VAR
END_METHOD

METHOD CALL_OUTPUT
END_METHOD

METHOD CALL_REQUESTS_EXT
END_METHOD

METHOD CALL_RESETCOMMANDS
END_METHOD

METHOD CALL_RESETOUTPUT
END_METHOD

METHOD CALL_STATEMACHINE
VAR_IN_OUT
	AXESGROUP : AXES_GROUP_KIN;
END_VAR
END_METHOD

METHOD CALL_UNLOCKPATHDATA
VAR_IN_OUT
	AXESGROUP : AXES_GROUP_KIN;
END_VAR
END_METHOD

METHOD FUN_ACKNLASTELEMENT : BOOL
VAR_INPUT
	PELEMENT : POINTER TO L_MC4P_Parameter_MCMove;
	IDX : INT;
END_VAR
END_METHOD

METHOD FUN_ACKNOWLEDGEELEMENT
VAR_INPUT
	IELEMENTNO : INT := 1;
END_VAR
END_METHOD

METHOD FUN_INITELEMENT
VAR_IN_OUT
	AXESGROUP : AXES_GROUP_KIN;
	SCPARELEMENT : L_MC4P_Parameter_MCMove;
END_VAR
END_METHOD

METHOD FUN_SEARCHFINALELEMENT : BOOL
END_METHOD

METHOD FB_INIT : BOOL
VAR_INPUT
	BINITRETAINS : BOOL;
	BINCOPYCODE : BOOL;
END_VAR
END_METHOD

METHOD CALL_PATHREFINFO
END_METHOD

METHOD CALL_INIT
END_METHOD

METHOD CALL_S000_CYCLIC
VAR_IN_OUT
	AXESGROUP : AXES_GROUP_KIN;
END_VAR
END_METHOD

(* ---- MC_READCARTESIANTRANSFORM.fb ---- *)
FUNCTION_BLOCK MC_READCARTESIANTRANSFORM EXTENDS L_MC4P_Template_AG_KIN
VAR_INPUT
	ENABLE : BOOL;
	COORDSYSTEM : L_MC4P_CoordSystem;
END_VAR
VAR_OUTPUT
	VALID : BOOL;
	BUSY : BOOL;
	ERROR : BOOL;
	ERRORID : L_IE1P_Error;
	TRANSX : LREAL;
	TRANSY : LREAL;
	TRANSZ : LREAL;
	ROTANGLE1 : LREAL;
	ROTANGLE2 : LREAL;
	ROTANGLE3 : LREAL;
END_VAR
VAR
	PCOORDTRAFO : POINTER TO L_MC4P_CoordTrafo;
	XENABLEOLD : BOOL;
END_VAR
END_FUNCTION_BLOCK

(* ---- MC_READCOORDINATETRANSFORM.fb ---- *)
FUNCTION_BLOCK MC_READCOORDINATETRANSFORM EXTENDS L_MC4P_Template_AG_KIN
VAR_INPUT
	ENABLE : BOOL;
	COORDSYSTEM : L_MC4P_CoordSystem;
END_VAR
VAR_OUTPUT
	VALID : BOOL;
	BUSY : BOOL;
	ERROR : BOOL;
	ERRORID : L_IE1P_Error;
	COORDTRANSFORM : MC_COORD_REF;
END_VAR
VAR
	PCOORDTRAFO : POINTER TO L_MC4P_CoordTrafo;
	XENABLEOLD : BOOL;
END_VAR
END_FUNCTION_BLOCK

(* ---- MC_REMOVEAXISFROMGROUP.fb ---- *)
FUNCTION_BLOCK MC_REMOVEAXISFROMGROUP EXTENDS L_MC4P_Template_AG_KIN
VAR_INPUT
	EXECUTE : BOOL;
	IDENTINGROUP : IDENT_IN_GROUP_REF;
END_VAR
VAR_OUTPUT
	DONE : BOOL;
	BUSY : BOOL;
	ERROR : BOOL;
	ERRORID : L_IE1P_Error;
END_VAR
VAR
	XERRORINTERN : BOOL;
	EERRORIDINTERN : L_IE1P_Error := L_IE1P_Error.NoError;
	XEXECUTEOLD : BOOL;
	XRESETOUTPUT : BOOL;
	PSDUMMY : POINTER TO STRING;
	DWINTERNALERRORID : DWORD;
END_VAR
END_FUNCTION_BLOCK

(* ---- MC_SETCARTESIANTRANSFORM.fb ---- *)
FUNCTION_BLOCK MC_SETCARTESIANTRANSFORM EXTENDS L_MC4P_Template_AG_KIN
VAR_INPUT
	EXECUTE : BOOL;
	COORDSYSTEM : L_MC4P_CoordSystem;
	TRANSX : LREAL;
	TRANSY : LREAL;
	TRANSZ : LREAL;
	ROTANGLE1 : LREAL;
	ROTANGLE2 : LREAL;
	ROTANGLE3 : LREAL;
END_VAR
VAR_OUTPUT
	DONE : BOOL;
	BUSY : BOOL;
	ACTIVE : BOOL;
	COMMANDABORTED : BOOL;
	ERROR : BOOL;
	ERRORID : L_IE1P_Error;
END_VAR
VAR
	PCOORDTRAFO : POINTER TO L_MC4P_CoordTrafo;
	XEXECUTEOLD : BOOL;
	XRESETOUTPUT : BOOL;
	ISTATE : INT;
	BSTATEMACHINE : BOOL;
	PTRACKINGPARAM : POINTER TO L_MC4P_PCSTrackParam;
	ALRPARAMFREEZE : ARRAY [1..6] OF LREAL;
	AXPARACCESSIBLE : ARRAY [1..7] OF BOOL;
	IDX : DINT;
	XINTERNALTESTMODE : BOOL := FALSE;
	INTERNALTESTMODE : BOOL;
END_VAR
END_FUNCTION_BLOCK

(* ---- MC_SETCOORDINATETRANSFORM.fb ---- *)
FUNCTION_BLOCK MC_SETCOORDINATETRANSFORM EXTENDS L_MC4P_Template_AG_KIN
VAR_INPUT
	EXECUTE : BOOL;
	COORDTRANSFORM : MC_COORD_REF;
	COORDSYSTEM : L_MC4P_CoordSystem;
END_VAR
VAR_OUTPUT
	DONE : BOOL;
	BUSY : BOOL;
	ACTIVE : BOOL;
	COMMANDABORTED : BOOL;
	ERROR : BOOL;
	ERRORID : L_IE1P_Error;
END_VAR
VAR
	PCOORDTRAFO : POINTER TO L_MC4P_CoordTrafo;
	XEXECUTEOLD : BOOL;
	XRESETOUTPUT : BOOL;
	ISTATE : INT;
	BSTATEMACHINE : BOOL;
	PTRACKINGPARAM : POINTER TO L_MC4P_PCSTrackParam;
	COORDTRANSFFREEZE : MC_COORD_REF;
	AXPARACCESSIBLE : ARRAY [1..7] OF BOOL;
	IDX : DINT;
	XINTERNALTESTMODE : BOOL := FALSE;
	INTERNALTESTMODE : BOOL;
END_VAR
END_FUNCTION_BLOCK

(* ---- MC_SETKINTRANSFORM.fb ---- *)
FUNCTION_BLOCK MC_SETKINTRANSFORM EXTENDS L_MC4P_Template_AG_KIN
VAR_INPUT
	EXECUTE : BOOL;
	KINTRANSFORM : MC_KIN_REF;
END_VAR
VAR_OUTPUT
	DONE : BOOL;
	BUSY : BOOL;
	ACTIVE : BOOL;
	COMMANDABORTED : BOOL;
	ERROR : BOOL;
	ERRORID : L_IE1P_Error;
END_VAR
VAR
	XEXECUTEOLD : BOOL;
	XRESETOUTPUT : BOOL;
	PAXESGROUP : POINTER TO AXES_GROUP_KIN;
END_VAR
END_FUNCTION_BLOCK

(* ---- MC_TRACKCONVEYORBELT.fb ---- *)
FUNCTION_BLOCK MC_TRACKCONVEYORBELT EXTENDS L_MC4P_Template_AG_KIN_Licence
VAR_INPUT
	EXECUTE : BOOL;
	ABORT : BOOL;
	CONVEYORBELTORIGIN : ARRAY [1..6] OF LREAL;
	INITIALOBJECTPOSITION : ARRAY [1..6] OF LREAL;
	COORDSYSTEM : L_MC4P_CoordSystem;
	COORDTYPE : L_MC4P_CoordType;
	CLUTCHDISTANCE : LREAL;
	CLUTCHTIME : LREAL;
	CLUTCHTIMEABORT : LREAL;
	SETDYNPCS : BOOL := TRUE;
END_VAR
VAR_OUTPUT
	DONE : BOOL;
	BUSY : BOOL;
	ACTIVE : BOOL;
	COMMANDABORTED : BOOL;
	ERROR : BOOL;
	ERRORID : L_IE1P_Error;
	INSYNC : BOOL;
	DYNAMICPCSSET : BOOL;
END_VAR
VAR_IN_OUT
	CONVEYORBELT : AXIS_REF;
END_VAR
VAR
	TRACK : L_MC4P_TrackConveyorBelt_internal;
	CLUTCHEXTERNAL : LREAL;
	MASTERVALUESOURCE : MC_SOURCE;
END_VAR
END_FUNCTION_BLOCK

(* ---- MC_UNGROUPALLAXES.fb ---- *)
FUNCTION_BLOCK MC_UNGROUPALLAXES EXTENDS L_MC4P_Template_AG_KIN
VAR_INPUT
	EXECUTE : BOOL;
END_VAR
VAR_OUTPUT
	DONE : BOOL;
	BUSY : BOOL;
	ERROR : BOOL;
	ERRORID : L_IE1P_Error;
END_VAR
VAR
	XEXECUTEOLD : BOOL;
	XRESETOUTPUT : BOOL;
	PSDUMMY : POINTER TO STRING;
	IDX : WORD;
END_VAR
END_FUNCTION_BLOCK
